      CALL "SENSOR CHECK" (
           Bit                      := "B 7.4",
           Preset_ms                := 500,
           Plc_Scan_ms              := "DB UTILITY".Scan_Cycle_Previous,
           Rising_Pulse_1           := "DB SENSOR CHECK".B7_4.Rising_Pulse_1,
           Rising_Pulse_2           := "DB SENSOR CHECK".B7_4.Rising_Pulse_2,
           Memory_Bit_1             := "DB SENSOR CHECK".B7_4.Memory_Bit_1,
           Memory_Bit_2             := "DB SENSOR CHECK".B7_4.Memory_Bit_2,
           Word_Buffer              := "DB SENSOR CHECK".B7_4.Word_buffer,
           Word_Result              := "DB SENSOR CHECK".B7_4.Word_Result);

NETWORK
TITLE =
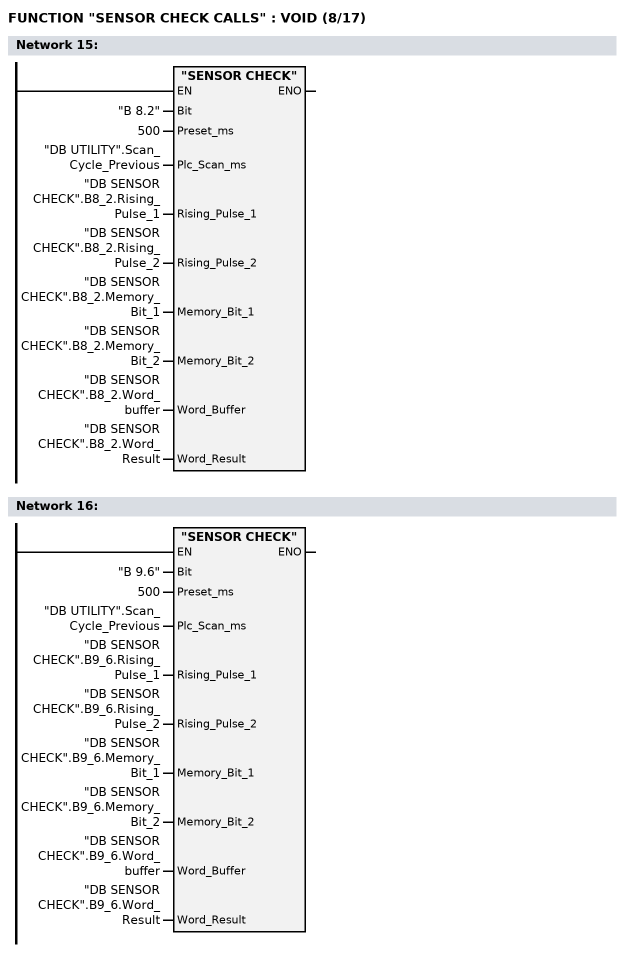

      CALL "SENSOR CHECK" (
           Bit                      := "B 8.2",
           Preset_ms                := 500,
           Plc_Scan_ms              := "DB UTILITY".Scan_Cycle_Previous,
           Rising_Pulse_1           := "DB SENSOR CHECK".B8_2.Rising_Pulse_1,
           Rising_Pulse_2           := "DB SENSOR CHECK".B8_2.Rising_Pulse_2,
           Memory_Bit_1             := "DB SENSOR CHECK".B8_2.Memory_Bit_1,
           Memory_Bit_2             := "DB SENSOR CHECK".B8_2.Memory_Bit_2,
           Word_Buffer              := "DB SENSOR CHECK".B8_2.Word_buffer,
           Word_Result              := "DB SENSOR CHECK".B8_2.Word_Result);

NETWORK
TITLE =

      CALL "SENSOR CHECK" (
           Bit                      := "B 9.6",
           Preset_ms                := 500,
           Plc_Scan_ms              := "DB UTILITY".Scan_Cycle_Previous,
           Rising_Pulse_1           := "DB SENSOR CHECK".B9_6.Rising_Pulse_1,
           Rising_Pulse_2           := "DB SENSOR CHECK".B9_6.Rising_Pulse_2,
           Memory_Bit_1             := "DB SENSOR CHECK".B9_6.Memory_Bit_1,
           Memory_Bit_2             := "DB SENSOR CHECK".B9_6.Memory_Bit_2,
           Word_Buffer              := "DB SENSOR CHECK".B9_6.Word_buffer,
           Word_Result              := "DB SENSOR CHECK".B9_6.Word_Result);

NETWORK
TITLE =
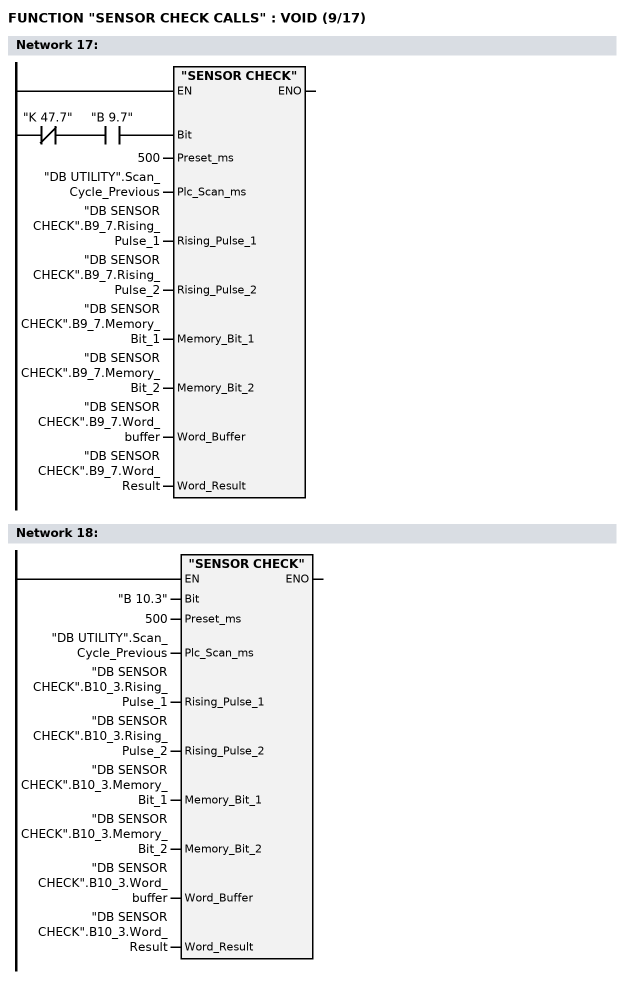

      AN    "K 47.7";
      A     "B 9.7";
      =     L      0.1;
//;
      CALL "SENSOR CHECK" (
           Bit                      := L      0.1,
           Preset_ms                := 500,
           Plc_Scan_ms              := "DB UTILITY".Scan_Cycle_Previous,
           Rising_Pulse_1           := "DB SENSOR CHECK".B9_7.Rising_Pulse_1,
           Rising_Pulse_2           := "DB SENSOR CHECK".B9_7.Rising_Pulse_2,
           Memory_Bit_1             := "DB SENSOR CHECK".B9_7.Memory_Bit_1,
           Memory_Bit_2             := "DB SENSOR CHECK".B9_7.Memory_Bit_2,
           Word_Buffer              := "DB SENSOR CHECK".B9_7.Word_buffer,
           Word_Result              := "DB SENSOR CHECK".B9_7.Word_Result);

NETWORK
TITLE =

      CALL "SENSOR CHECK" (
           Bit                      := "B 10.3",
           Preset_ms                := 500,
           Plc_Scan_ms              := "DB UTILITY".Scan_Cycle_Previous,
           Rising_Pulse_1           := "DB SENSOR CHECK".B10_3.Rising_Pulse_1,
           Rising_Pulse_2           := "DB SENSOR CHECK".B10_3.Rising_Pulse_2,
           Memory_Bit_1             := "DB SENSOR CHECK".B10_3.Memory_Bit_1,
           Memory_Bit_2             := "DB SENSOR CHECK".B10_3.Memory_Bit_2,
           Word_Buffer              := "DB SENSOR CHECK".B10_3.Word_buffer,
           Word_Result              := "DB SENSOR CHECK".B10_3.Word_Result);

NETWORK
TITLE =
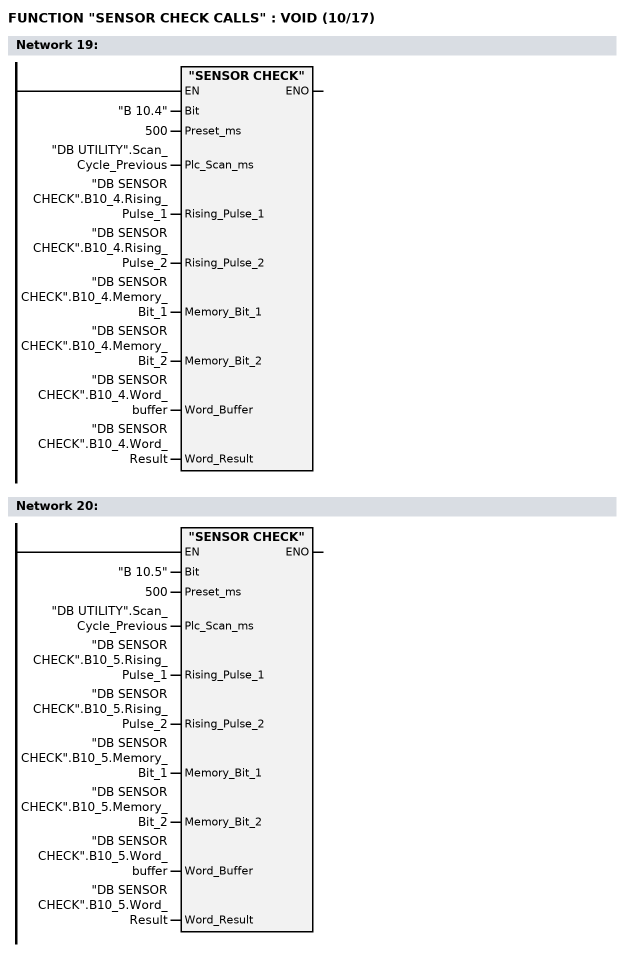

      CALL "SENSOR CHECK" (
           Bit                      := "B 10.4",
           Preset_ms                := 500,
           Plc_Scan_ms              := "DB UTILITY".Scan_Cycle_Previous,
           Rising_Pulse_1           := "DB SENSOR CHECK".B10_4.Rising_Pulse_1,
           Rising_Pulse_2           := "DB SENSOR CHECK".B10_4.Rising_Pulse_2,
           Memory_Bit_1             := "DB SENSOR CHECK".B10_4.Memory_Bit_1,
           Memory_Bit_2             := "DB SENSOR CHECK".B10_4.Memory_Bit_2,
           Word_Buffer              := "DB SENSOR CHECK".B10_4.Word_buffer,
           Word_Result              := "DB SENSOR CHECK".B10_4.Word_Result);

NETWORK
TITLE =

      CALL "SENSOR CHECK" (
           Bit                      := "B 10.5",
           Preset_ms                := 500,
           Plc_Scan_ms              := "DB UTILITY".Scan_Cycle_Previous,
           Rising_Pulse_1           := "DB SENSOR CHECK".B10_5.Rising_Pulse_1,
           Rising_Pulse_2           := "DB SENSOR CHECK".B10_5.Rising_Pulse_2,
           Memory_Bit_1             := "DB SENSOR CHECK".B10_5.Memory_Bit_1,
           Memory_Bit_2             := "DB SENSOR CHECK".B10_5.Memory_Bit_2,
           Word_Buffer              := "DB SENSOR CHECK".B10_5.Word_buffer,
           Word_Result              := "DB SENSOR CHECK".B10_5.Word_Result);

NETWORK
TITLE =
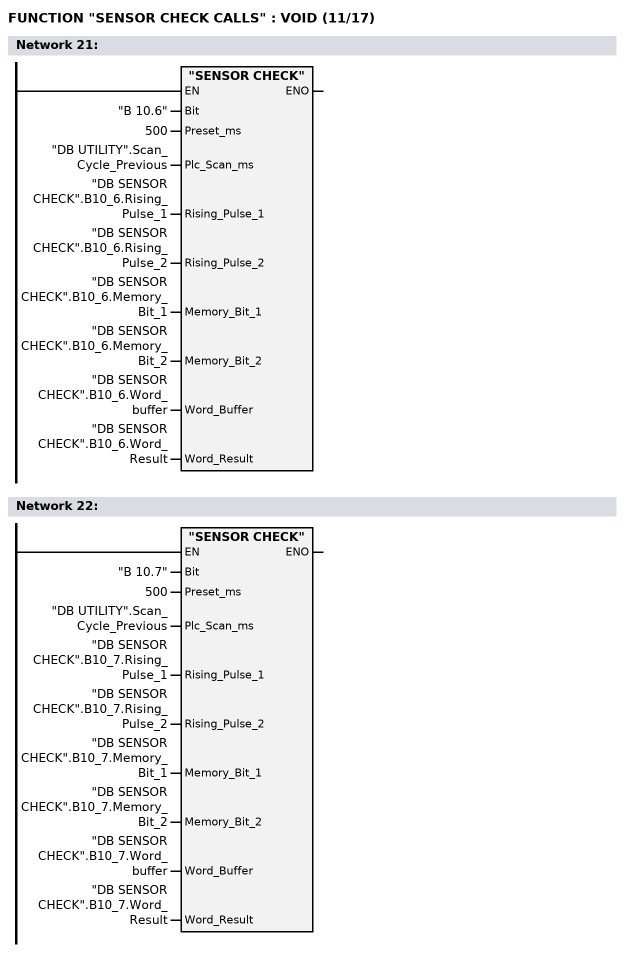

      CALL "SENSOR CHECK" (
           Bit                      := "B 10.6",
           Preset_ms                := 500,
           Plc_Scan_ms              := "DB UTILITY".Scan_Cycle_Previous,
           Rising_Pulse_1           := "DB SENSOR CHECK".B10_6.Rising_Pulse_1,
           Rising_Pulse_2           := "DB SENSOR CHECK".B10_6.Rising_Pulse_2,
           Memory_Bit_1             := "DB SENSOR CHECK".B10_6.Memory_Bit_1,
           Memory_Bit_2             := "DB SENSOR CHECK".B10_6.Memory_Bit_2,
           Word_Buffer              := "DB SENSOR CHECK".B10_6.Word_buffer,
           Word_Result              := "DB SENSOR CHECK".B10_6.Word_Result);

NETWORK
TITLE =

      CALL "SENSOR CHECK" (
           Bit                      := "B 10.7",
           Preset_ms                := 500,
           Plc_Scan_ms              := "DB UTILITY".Scan_Cycle_Previous,
           Rising_Pulse_1           := "DB SENSOR CHECK".B10_7.Rising_Pulse_1,
           Rising_Pulse_2           := "DB SENSOR CHECK".B10_7.Rising_Pulse_2,
           Memory_Bit_1             := "DB SENSOR CHECK".B10_7.Memory_Bit_1,
           Memory_Bit_2             := "DB SENSOR CHECK".B10_7.Memory_Bit_2,
           Word_Buffer              := "DB SENSOR CHECK".B10_7.Word_buffer,
           Word_Result              := "DB SENSOR CHECK".B10_7.Word_Result);

NETWORK
TITLE =
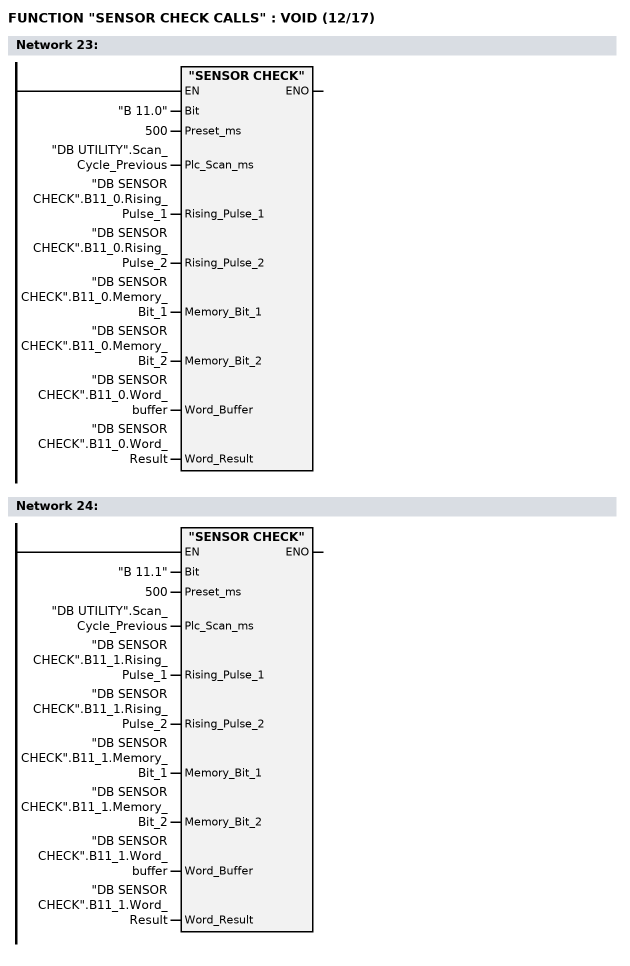

      CALL "SENSOR CHECK" (
           Bit                      := "B 11.0",
           Preset_ms                := 500,
           Plc_Scan_ms              := "DB UTILITY".Scan_Cycle_Previous,
           Rising_Pulse_1           := "DB SENSOR CHECK".B11_0.Rising_Pulse_1,
           Rising_Pulse_2           := "DB SENSOR CHECK".B11_0.Rising_Pulse_2,
           Memory_Bit_1             := "DB SENSOR CHECK".B11_0.Memory_Bit_1,
           Memory_Bit_2             := "DB SENSOR CHECK".B11_0.Memory_Bit_2,
           Word_Buffer              := "DB SENSOR CHECK".B11_0.Word_buffer,
           Word_Result              := "DB SENSOR CHECK".B11_0.Word_Result);

NETWORK
TITLE =

      CALL "SENSOR CHECK" (
           Bit                      := "B 11.1",
           Preset_ms                := 500,
           Plc_Scan_ms              := "DB UTILITY".Scan_Cycle_Previous,
           Rising_Pulse_1           := "DB SENSOR CHECK".B11_1.Rising_Pulse_1,
           Rising_Pulse_2           := "DB SENSOR CHECK".B11_1.Rising_Pulse_2,
           Memory_Bit_1             := "DB SENSOR CHECK".B11_1.Memory_Bit_1,
           Memory_Bit_2             := "DB SENSOR CHECK".B11_1.Memory_Bit_2,
           Word_Buffer              := "DB SENSOR CHECK".B11_1.Word_buffer,
           Word_Result              := "DB SENSOR CHECK".B11_1.Word_Result);

NETWORK
TITLE =
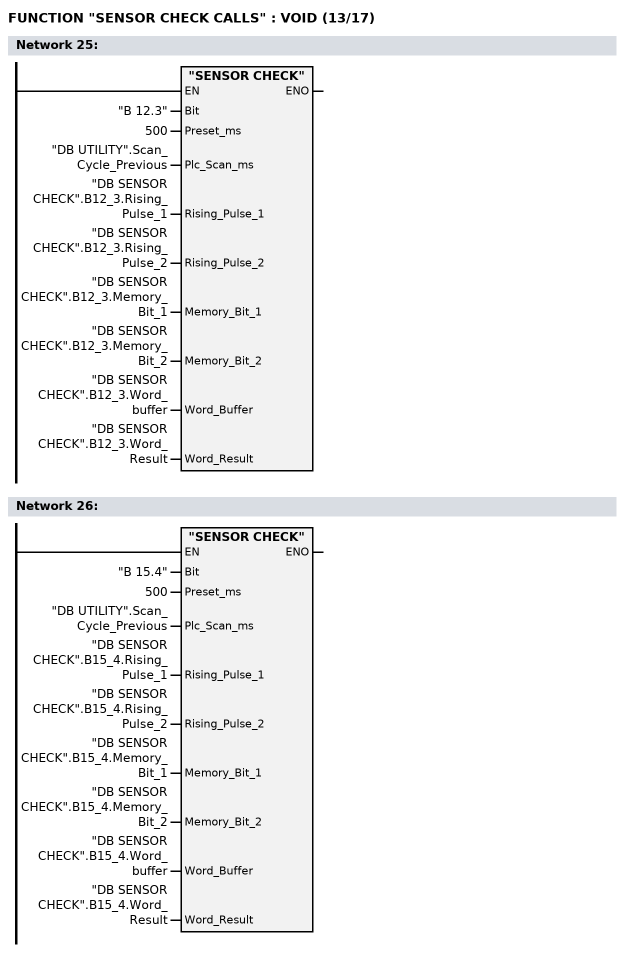

      CALL "SENSOR CHECK" (
           Bit                      := "B 12.3",
           Preset_ms                := 500,
           Plc_Scan_ms              := "DB UTILITY".Scan_Cycle_Previous,
           Rising_Pulse_1           := "DB SENSOR CHECK".B12_3.Rising_Pulse_1,
           Rising_Pulse_2           := "DB SENSOR CHECK".B12_3.Rising_Pulse_2,
           Memory_Bit_1             := "DB SENSOR CHECK".B12_3.Memory_Bit_1,
           Memory_Bit_2             := "DB SENSOR CHECK".B12_3.Memory_Bit_2,
           Word_Buffer              := "DB SENSOR CHECK".B12_3.Word_buffer,
           Word_Result              := "DB SENSOR CHECK".B12_3.Word_Result);

NETWORK
TITLE =

      CALL "SENSOR CHECK" (
           Bit                      := "B 15.4",
           Preset_ms                := 500,
           Plc_Scan_ms              := "DB UTILITY".Scan_Cycle_Previous,
           Rising_Pulse_1           := "DB SENSOR CHECK".B15_4.Rising_Pulse_1,
           Rising_Pulse_2           := "DB SENSOR CHECK".B15_4.Rising_Pulse_2,
           Memory_Bit_1             := "DB SENSOR CHECK".B15_4.Memory_Bit_1,
           Memory_Bit_2             := "DB SENSOR CHECK".B15_4.Memory_Bit_2,
           Word_Buffer              := "DB SENSOR CHECK".B15_4.Word_buffer,
           Word_Result              := "DB SENSOR CHECK".B15_4.Word_Result);

NETWORK
TITLE =
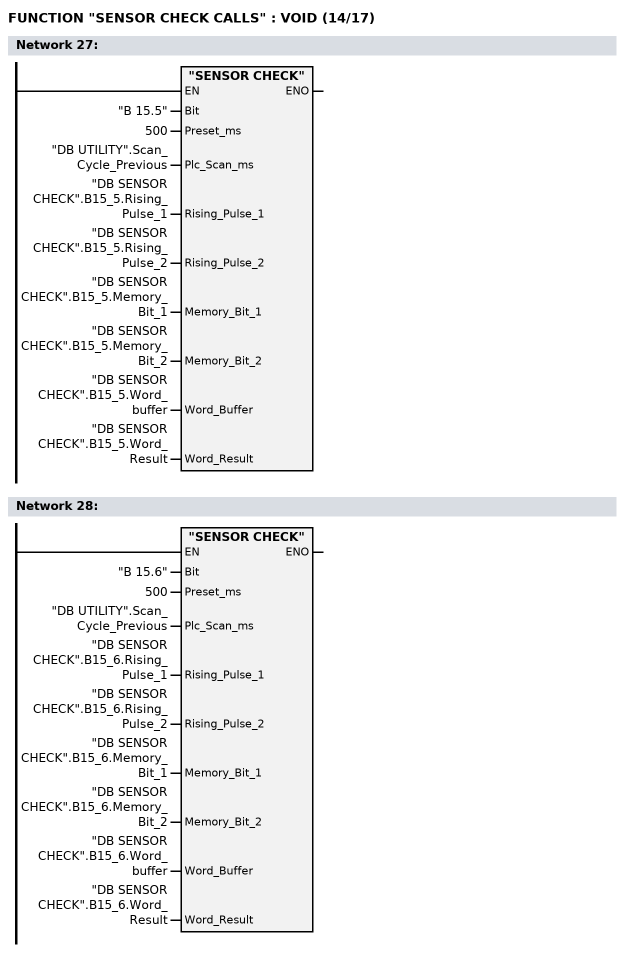

      CALL "SENSOR CHECK" (
           Bit                      := "B 15.5",
           Preset_ms                := 500,
           Plc_Scan_ms              := "DB UTILITY".Scan_Cycle_Previous,
           Rising_Pulse_1           := "DB SENSOR CHECK".B15_5.Rising_Pulse_1,
           Rising_Pulse_2           := "DB SENSOR CHECK".B15_5.Rising_Pulse_2,
           Memory_Bit_1             := "DB SENSOR CHECK".B15_5.Memory_Bit_1,
           Memory_Bit_2             := "DB SENSOR CHECK".B15_5.Memory_Bit_2,
           Word_Buffer              := "DB SENSOR CHECK".B15_5.Word_buffer,
           Word_Result              := "DB SENSOR CHECK".B15_5.Word_Result);

NETWORK
TITLE =

      CALL "SENSOR CHECK" (
           Bit                      := "B 15.6",
           Preset_ms                := 500,
           Plc_Scan_ms              := "DB UTILITY".Scan_Cycle_Previous,
           Rising_Pulse_1           := "DB SENSOR CHECK".B15_6.Rising_Pulse_1,
           Rising_Pulse_2           := "DB SENSOR CHECK".B15_6.Rising_Pulse_2,
           Memory_Bit_1             := "DB SENSOR CHECK".B15_6.Memory_Bit_1,
           Memory_Bit_2             := "DB SENSOR CHECK".B15_6.Memory_Bit_2,
           Word_Buffer              := "DB SENSOR CHECK".B15_6.Word_buffer,
           Word_Result              := "DB SENSOR CHECK".B15_6.Word_Result);

NETWORK
TITLE =
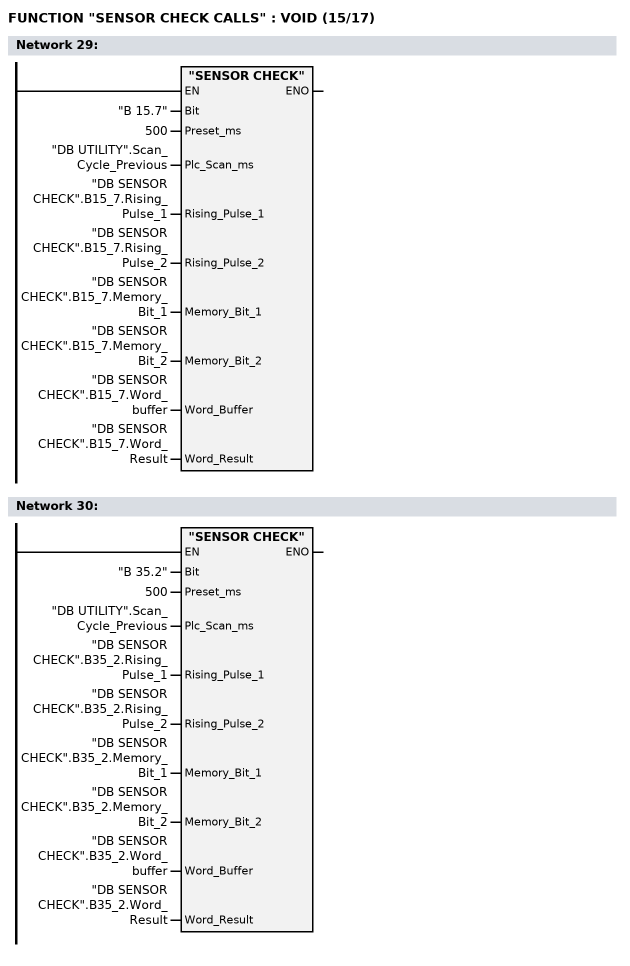

      CALL "SENSOR CHECK" (
           Bit                      := "B 15.7",
           Preset_ms                := 500,
           Plc_Scan_ms              := "DB UTILITY".Scan_Cycle_Previous,
           Rising_Pulse_1           := "DB SENSOR CHECK".B15_7.Rising_Pulse_1,
           Rising_Pulse_2           := "DB SENSOR CHECK".B15_7.Rising_Pulse_2,
           Memory_Bit_1             := "DB SENSOR CHECK".B15_7.Memory_Bit_1,
           Memory_Bit_2             := "DB SENSOR CHECK".B15_7.Memory_Bit_2,
           Word_Buffer              := "DB SENSOR CHECK".B15_7.Word_buffer,
           Word_Result              := "DB SENSOR CHECK".B15_7.Word_Result);

NETWORK
TITLE =

      CALL "SENSOR CHECK" (
           Bit                      := "B 35.2",
           Preset_ms                := 500,
           Plc_Scan_ms              := "DB UTILITY".Scan_Cycle_Previous,
           Rising_Pulse_1           := "DB SENSOR CHECK".B35_2.Rising_Pulse_1,
           Rising_Pulse_2           := "DB SENSOR CHECK".B35_2.Rising_Pulse_2,
           Memory_Bit_1             := "DB SENSOR CHECK".B35_2.Memory_Bit_1,
           Memory_Bit_2             := "DB SENSOR CHECK".B35_2.Memory_Bit_2,
           Word_Buffer              := "DB SENSOR CHECK".B35_2.Word_buffer,
           Word_Result              := "DB SENSOR CHECK".B35_2.Word_Result);

NETWORK
TITLE =
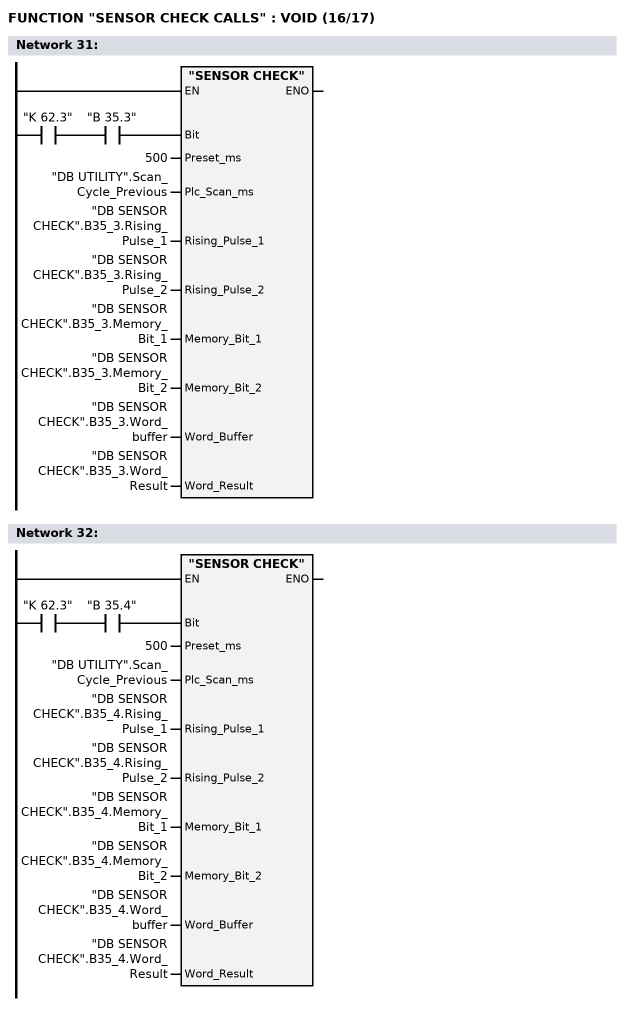

      A     "K 62.3";
      A     "B 35.3";
      =     L      0.2;

      CALL "SENSOR CHECK" (
           Bit                      := L      0.2,
           Preset_ms                := 500,
           Plc_Scan_ms              := "DB UTILITY".Scan_Cycle_Previous,
           Rising_Pulse_1           := "DB SENSOR CHECK".B35_3.Rising_Pulse_1,
           Rising_Pulse_2           := "DB SENSOR CHECK".B35_3.Rising_Pulse_2,
           Memory_Bit_1             := "DB SENSOR CHECK".B35_3.Memory_Bit_1,
           Memory_Bit_2             := "DB SENSOR CHECK".B35_3.Memory_Bit_2,
           Word_Buffer              := "DB SENSOR CHECK".B35_3.Word_buffer,
           Word_Result              := "DB SENSOR CHECK".B35_3.Word_Result);

NETWORK
TITLE =

      A     "K 62.3";
      A     "B 35.4";
      =     L      0.3;
//;
      CALL "SENSOR CHECK" (
           Bit                      := L      0.3,
           Preset_ms                := 500,
           Plc_Scan_ms              := "DB UTILITY".Scan_Cycle_Previous,
           Rising_Pulse_1           := "DB SENSOR CHECK".B35_4.Rising_Pulse_1,
           Rising_Pulse_2           := "DB SENSOR CHECK".B35_4.Rising_Pulse_2,
           Memory_Bit_1             := "DB SENSOR CHECK".B35_4.Memory_Bit_1,
           Memory_Bit_2             := "DB SENSOR CHECK".B35_4.Memory_Bit_2,
           Word_Buffer              := "DB SENSOR CHECK".B35_4.Word_buffer,
           Word_Result              := "DB SENSOR CHECK".B35_4.Word_Result);

NETWORK
TITLE =
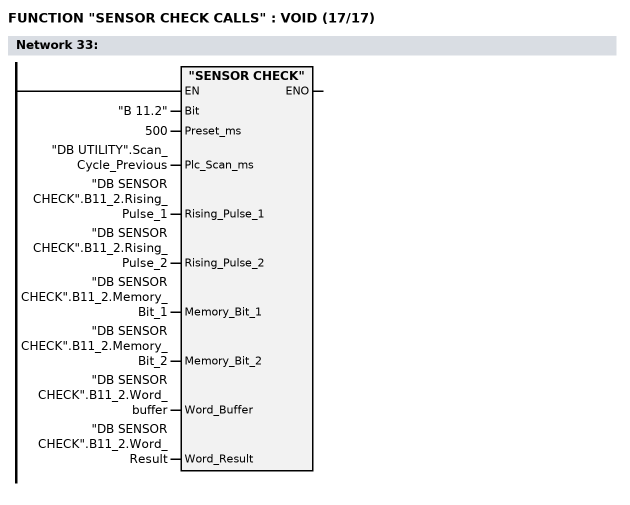

      CALL "SENSOR CHECK" (
           Bit                      := "B 11.2",
           Preset_ms                := 500,
           Plc_Scan_ms              := "DB UTILITY".Scan_Cycle_Previous,
           Rising_Pulse_1           := "DB SENSOR CHECK".B11_2.Rising_Pulse_1,
           Rising_Pulse_2           := "DB SENSOR CHECK".B11_2.Rising_Pulse_2,
           Memory_Bit_1             := "DB SENSOR CHECK".B11_2.Memory_Bit_1,
           Memory_Bit_2             := "DB SENSOR CHECK".B11_2.Memory_Bit_2,
           Word_Buffer              := "DB SENSOR CHECK".B11_2.Word_buffer,
           Word_Result              := "DB SENSOR CHECK".B11_2.Word_Result);

END_FUNCTION

FUNCTION "LAUER_RE-START_PUP" : VOID
TITLE =
//Logique de remise à zéro du bit de redémarrage de la communication avec
//l'interface.
//
//Ce bit doit être remis à zéro en cas de perte de communication avec l'automate
//ou si l'interface est éteint.
VERSION : 0.1

BEGIN
NETWORK
TITLE =Lauer restart bit
//DB50.DBW25 = S and mS   “Start a 5-second watchdog timer unless reset is
//active”
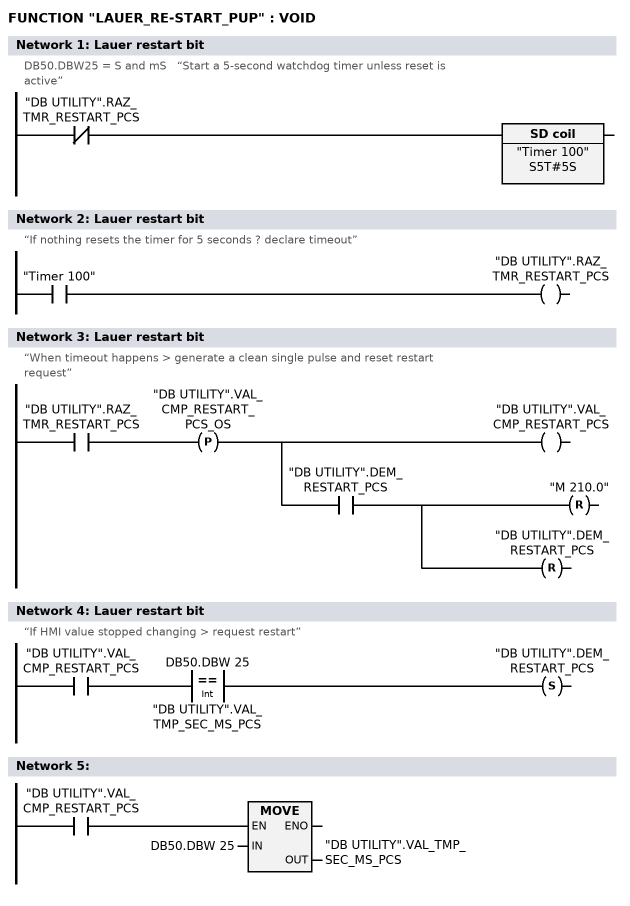
      AN    "DB UTILITY".RAZ_TMR_RESTART_PCS;
      L     S5T#5S;
      SD    "Timer 100";
      NOP   0;
      NOP   0;
      NOP   0;
      NOP   0;
NETWORK
TITLE =Lauer restart bit
//“If nothing resets the timer for 5 seconds ? declare timeout”
      A     "Timer 100";
      =     "DB UTILITY".RAZ_TMR_RESTART_PCS;
NETWORK
TITLE =Lauer restart bit
//“When timeout happens > generate a clean single pulse and reset restart
//request”
      A     "DB UTILITY".RAZ_TMR_RESTART_PCS;
      FP    "DB UTILITY".VAL_CMP_RESTART_PCS_OS;
      =     L      0.0;
      A     L      0.0;
      BLD   102;
      =     "DB UTILITY".VAL_CMP_RESTART_PCS;
      A     L      0.0;
      A     "DB UTILITY".DEM_RESTART_PCS;
      R     "M 210.0";
      R     "DB UTILITY".DEM_RESTART_PCS;
NETWORK
TITLE =Lauer restart bit
//“If HMI value stopped changing > request restart”
      A     "DB UTILITY".VAL_CMP_RESTART_PCS;
      A(    ;
      L     DB50.DBW   25;
      L     "DB UTILITY".VAL_TMP_SEC_MS_PCS;
      ==I   ;
      )     ;
      S     "DB UTILITY".DEM_RESTART_PCS;
NETWORK
TITLE =

      A     "DB UTILITY".VAL_CMP_RESTART_PCS;
      JNB   _001;
      L     DB50.DBW   25;
      T     "DB UTILITY".VAL_TMP_SEC_MS_PCS;
_001: NOP   0;
END_FUNCTION

FUNCTION "LAUER COMM ERR FC" : VOID
TITLE =
VERSION : 0.1

BEGIN
NETWORK
TITLE =
//;    Please choose your PCS and add the commands to your network
//;                      // Example PCS900/PCS 920/PCS950
//;                      // Typical presets
//;L W#16#1F00;  //(3F00 PCS950/PCS 920)
//;T DBW 72;
//;L W#16#00FF;
//;T DBW 74;
//;L W#16#0080;
//:T DBW 76;
//;                      // Example PCS009/PCS090/PCS095
//;                      // Typical presets
//;     L W#16#0FC8;
//;     T DBW 26;
//;     L W#16#0080;
//;     T DBW 28;
      L     W#16#0;
      T     DBW    8;
      T     DBW   10;
      T     DBW   12;
      T     DBW   14;
      T     DBW   46;
END_FUNCTION

FUNCTION "LAUER RESTART FC" : VOID
TITLE =
NAME : COFF
VERSION : 0.0

BEGIN
NETWORK
TITLE =
//;                     // Presets emergancy case
//;// Clear all keys
      L     W#16#0;
      T     DBW    8;
      T     DBW   10;
      T     DBW   12;
      T     DBW   14;
      T     DBW   46;
END_FUNCTION

FUNCTION "LAUER COMM FC" : VOID
TITLE =Handling Block Profibus
//
NAME : PROFIBUS
VERSION : 0.0


VAR_INPUT
  UBDB : BLOCK_DB ;	// UBDB
  RXFA : INT ;	// RXFA
  RXLE : INT ;	// RXLE
  TXFA : INT ;	// TXFA
  TXLE : INT ;	// TXLE
  RSET : BOOL ;	// RSET
  TIMT : TIMER ;	// TIMT
  TIMZ : S5TIME ;	// TIMZ
  COFF : BLOCK_FC ;	// COFF
  INIT : BLOCK_FC ;	// INIT
END_VAR
VAR_OUTPUT
  RFLM : BOOL ;	// RFLM
  EROR : BOOL ;	// EROR
END_VAR
VAR_TEMP
  conv_akku1 : DWORD ;
  conv_akku2 : DWORD ;
  conv_stw : WORD ;
END_VAR
BEGIN
NETWORK
TITLE =

      OPN   #UBDB; //  --------------------------
      AN    #RFLM; //  First action in FB?
      JC    OK;
      A     #TIMT; //  Timeout and no restart?
      AN    #RSET;
      JC    ERR;
      A     #TIMT;
      AN    #EROR;
      JC    ERR;
      JU    OK;

ERR:  A     #EROR;
      JC    ERR1;
      UC    #COFF; //  Call COFF once.
      OPN   #UBDB;

ERR1: A     #TIMT; //  If timeout set error-flag.
      S     #EROR;
      BEU   ;

OK:   A     #RFLM; //  First action?
      JC    CONT;
      UC    #INIT; //  Call INIT once.
      OPN   #UBDB;
      L     W#16#0; //  Init ----------------------
      T     DBW    0;
      T     DBW    2;
      T     DBW    4;
      T     DBW    6;
      AN    #RFLM;
      S     #RFLM; //  Set reset-ready-flag
//;
      AN    #RFLM; //  Trigger timer
      L     #TIMZ;
      SD    #TIMT;
//;
      A     #RFLM;
      L     #TIMZ;
      SD    #TIMT;

CONT: L     #RXFA;
      T     "MW 244"; //  ----------------------------
      +     1; //  Adress Handle1 E-Box
      T     "MW 252";
      L     #RXLE; //  Adress of first instruction
      +     -2;
      T     "MW 250"; //  Lenght E-Box Userdatas
//;
      L     #TXFA;
      T     "MW 242";
      +     1; //  Adress Handle1 A-Box
      T     "MW 248";
      L     #TXLE; //  Adress of first senddata
      +     -2;
      T     "MW 246"; //  Lenght A-Box-Userdatas
//;
      L     "MW 244"; //  Handle2 != Handle1? ---------
      L     #RXLE;
      +I    ;
      +     -1;
      T     "MW 238"; //  Adress Handle2
      T     #conv_akku1;
//;
      L     STW;
      T     #conv_stw;
//;
      L     "MB 239";
      SLW   3;
      LAR1  ;
      L     #conv_stw;
      T     STW;
//;
      L     #conv_akku1;
      L     IB [AR1,P#0.0];
      T     "MW 238"; //  Handle2
      T     #conv_akku1; //  Adress Handle1
//;
      L     STW;
      T     #conv_stw;
//;
      L     "MB 245";
      SLW   3;
      LAR1  ;
      L     #conv_stw;
      T     STW;
//;
      L     #conv_akku1;
      L     IB [AR1,P#0.0];
      L     "MW 238";
      <>I   ;
      BEC   ; //  Handle1 != Handle2 -> EXIT
//;
      T     #conv_akku1; //  Handle1 != HandleAlt? -------

      L     STW;
      T     #conv_stw;
//;
      L     "MB 245";
      SLW   3;
      LAR1  ;
      L     #conv_stw;
      T     STW;
//;
      L     #conv_akku1;
      L     IB [AR1,P#0.0];
      L     DBW    0; //  HandleAlt in UBDB (0)
      ==I   ;
      BEC   ;
//;
      AN    #RFLM; //  Start timeout-timer
      L     #TIMZ;
      SD    #TIMT;
//;
      A     #RFLM;
      L     #TIMZ;
      SD    #TIMT;
//;
      T     #conv_akku1; //  First action requiered?
      L     STW;
      T     #conv_stw;
      L     "MB 245";
      SLW   3;
      LAR1  ;
      L     #conv_stw;
      T     STW;
//;
      L     #conv_akku1;
      L     IB [AR1,P#0.0];
      L     W#16#80; //  Handle == 0x80?
      <>I   ;
      JC    SLP1;
      A     #RSET; // Clear Restart-Flag.
      R     #RSET;

END:  NOP   0;

      T     #conv_akku1; // Get Handle1(E) from RX-Box.

      L     STW;
      T     #conv_stw;
//;
      L     "MB 245";
      SLW   3;
      LAR1  ;
      L     #conv_stw;
      T     STW;
//;
      L     #conv_akku1;
      L     IB [AR1,P#0.0];
      T     DBW    0; // Save to HandleAlt.
      INVI  ; // Invert.
      T     "MW 236"; // Temporary saved.
      L     "MW 236";
      T     #conv_akku1; // Take inverted Handle1(E) to
      TAK   ;
      T     #conv_akku2;
      L     STW;
      T     #conv_stw;
//;
      L     "MB 243";
      SLW   3;
      LAR1  ;
      L     #conv_stw;
      T     STW;
//;
      L     #conv_akku2;
      L     #conv_akku1;
      T     QB [AR1,P#0.0]; // Handle1(A).
//;
      L     "MW 242";
      L     #TXLE;
      +I    ;
      +     -1;
      T     "MW 238"; // Take inverted Handle1(E) to
      L     "MW 236";
      T     #conv_akku1;
      TAK   ;
      T     #conv_akku2;
      L     STW;
      T     #conv_stw;
//;
      L     "MB 239";
      SLW   3;
      LAR1  ;
      L     #conv_stw;
      T     STW;
//;
      L     #conv_akku2;
      L     #conv_akku1;
      T     QB [AR1,P#0.0];
//;
      AN    #TIMT; // Clear Error-Mark.
      R     #EROR;
      BEU   ; // see you later...

SLP1: L     #RXFA; // Reached Rx-Box-End?
      L     #RXLE;
      +I    ;
      +     -1;
      L     "MW 252";
      ==I   ;
      JC    END;

      T     #conv_akku1; //  Start/Continue--------------

      L     STW;
      T     #conv_stw;
//;
      L     "MB 253";
      SLW   3;
      LAR1  ;
      L     #conv_stw;
      T     STW;
//;
      L     #conv_akku1;
      L     IW [AR1,P#0.0];
      L     W#16#0; //  Is anything usable?
      ==I   ;
      JC    END;

      T     #conv_akku1; //  Get first ABW.

      L     STW;
      T     #conv_stw;
//;
      L     "MB 253";
      SLW   3;
      LAR1  ;
      L     #conv_stw;
      T     STW;
//;
      L     #conv_akku1;
      L     IB [AR1,P#0.0];
      T     "MW 240"; //  Adress(UBDB) in ABW.
      L     "MW 252";
      +     1; //  Increment RX-Pointer.
      T     "MW 252";
      T     #conv_akku1;
      L     STW;
      T     #conv_stw;
      L     "MB 253";
      SLW   3;
      LAR1  ;
      L     #conv_stw;
      T     STW;
//;
      L     #conv_akku1;
      L     IB [AR1,P#0.0]; //  Count of ABW: Bit3..0.
      T     "MW 238"; //  Command of ABW: Bit 7..4.
      L     "MW 252"; //  ABW pointer to next ABW
      +     1; //  or first data.
      T     "MW 252";
//;
      L     "MW 238"; //  Check for right command.
      L     W#16#F0;
      AW    ;
      T     "MW 236"; //  Temporary saved.
//;
      L     "MW 236";
      L     W#16#10;
      ==I   ;
      JC    IOK;
//;
      L     "MW 236";
      L     W#16#20;
      ==I   ;
      JC    IOK;
//;
      L     "MW 236";
      L     W#16#40;
      ==I   ;
      JC    IOK;
//;
      L     "MW 236";
      L     W#16#80;
      ==I   ;
      JC    IOK;
      BEU   ; //  Command is wrong!
//;
IOK:  L     "MW 238"; //  Command is ok.
SLP2: L     W#16#F;
      AW    ; //  Count == 0:
      JZ    SLP1; //  Next subpaket
//;
      AN    "M 239.4";
      JC    ELS1;
      OPN   #UBDB;

      T     #conv_akku1; //  Offset ABW Adress in UBDB

      L     STW;
      T     #conv_stw;
//;
      L     "MB 241";
      SLW   4;
      LAR1  ;
      L     #conv_stw;
      T     STW;
//;
      L     #conv_akku1;
      L     DBW [AR1,P#0.0];
      T     #conv_akku1; //  Pointer to TX-Box
      TAK   ;
      T     #conv_akku2;
      L     STW;
      T     #conv_stw;
//;
      L     "MB 249";
      SLW   3;
      LAR1  ;
      L     #conv_stw;
      T     STW;
//;
      L     #conv_akku2;
      L     #conv_akku1;
      T     QW [AR1,P#0.0]; //  Write to TX-Box.
      L     "MW 248";
      +     2;
      T     "MW 248";
      JU    COMM;

ELS1: NOP   0;

      T     #conv_akku1; //  Pointer to RX-Box.

      L     STW;
      T     #conv_stw;
//;
      L     "MB 253";
      SLW   3;
      LAR1  ;
      L     #conv_stw;
      T     STW;
//;
      L     #conv_akku1;
      L     IW [AR1,P#0.0];
      T     "MW 236"; //  Read Data/Mask from RX-Box.
      L     "MW 252"; //  Increment Pointer to RX-Box.
      +     2;
      T     "MW 252";
//;
      AN    "M 239.5"; //  WRITE/(AND/OR)
      JC    ELS2;
      L     "MW 236";
      OPN   #UBDB;

      T     #conv_akku1; //  Offset ABW Adress in UBDB.
      TAK   ;
      T     #conv_akku2;
      L     STW;
      T     #conv_stw;
      L     "MB 241";
      SLW   4;
      LAR1  ;
      L     #conv_stw;
      T     STW;
//;
      L     #conv_akku2;
      L     #conv_akku1;
      T     DBW [AR1,P#0.0]; //  Write to UBDB.
      JU    COMM;

ELS2: AN    "M 239.6";
      JC    ELS3;
      L     "MW 236";
      OPN   #UBDB;

      T     #conv_akku1; //  Offset ABW Adress in UBDB.
      L     STW;
      T     #conv_stw;
      L     "MB 241";
      SLW   4;
      LAR1  ;
      L     #conv_stw;
      T     STW;
//;
      L     #conv_akku1;
      L     DBW [AR1,P#0.0];
      AW    ;
      OPN   #UBDB;
      T     #conv_akku1;
      TAK   ;
      T     #conv_akku2;
      L     STW;
      T     #conv_stw;
      L     "MB 241";
      SLW   4;
      LAR1  ;
      L     #conv_stw;
      T     STW;
//;
      L     #conv_akku2;
      L     #conv_akku1;
      T     DBW [AR1,P#0.0]; //  And to UBDB
      JU    COMM;

ELS3: NOP   0;

      L     "MW 236";
      OPN   #UBDB;
      T     #conv_akku1;
      L     STW;
      T     #conv_stw;
      L     "MB 241";
      SLW   4;
      LAR1  ;
      L     #conv_stw;
      T     STW;
//;
      L     #conv_akku1;
      L     DBW [AR1,P#0.0];
      OW    ;
      OPN   #UBDB;

      T     #conv_akku1;
      TAK   ;
      T     #conv_akku2;
      L     STW;
      T     #conv_stw;
      L     "MB 241";
      SLW   4;
      LAR1  ;
      L     #conv_stw;
      T     STW;
//;
      L     #conv_akku2;
      L     #conv_akku1;
      T     DBW [AR1,P#0.0];
COMM: L     "MW 240";
      +     1;
      T     "MW 240";
      L     "MW 238"; //  Decrement counter of ABW.
      +     -1;
      T     "MW 238";
      JU    SLP2;
END_FUNCTION

FUNCTION "LAUER" : VOID
TITLE =
NAME : SCHRIANZ
VERSION : 0.0


VAR_TEMP
  TEMP0 : DWORD ;
  TEMP1 : DWORD ;
  TEMP2 : WORD ;
END_VAR
BEGIN
NETWORK
TITLE =



NETWORK
TITLE =



NETWORK
TITLE =

      OPN   "DB LAUER";

NETWORK
TITLE =

      AN    "M 150.7";
      JC    M001;
      L     2#100000000;
      T     DBW   72;
M001: NOP   0;
NETWORK
TITLE =

      ON    "M 150.7";
      JC    M002;
      L     2#1;
      T     DBW   76;
M002: NOP   0;
NETWORK
TITLE =



NETWORK
TITLE =

      O(    ;
      L     DBW  300;
      L     77;
      <I    ;
      )     ;
      O(    ;
      L     DBW  300;
      L     102;
      >I    ;
      )     ;
      JC    M003;
      JU    M004;
M003: L     77;
      T     DBW  300;
M004: NOP   0;
NETWORK
TITLE =

      L     "DB LAUER".D_150;
      L     77;
      <>I   ;
      JC    M005;
      L     "MW 15";
      T     "MW 200";
      L     "MB 17";
      T     MB   202;
M005: L     DBW  300;
      L     78;
      <>I   ;
      JC    M006;
      L     "MW 19";
      T     "MW 200";
      L     "MB 21";
      T     MB   202;
M006: L     DBW  300;
      L     79;
      <>I   ;
      JC    M007;
      L     "MW 23";
      T     "MW 200";
      L     "MB 25";
      T     MB   202;
M007: L     DBW  300;
      L     80;
      <>I   ;
      JC    M008;
      L     "MW 27";
      T     "MW 200";
      L     "MB 29";
      T     MB   202;
M008: L     DBW  300;
      L     81;
      <>I   ;
      JC    M009;
      L     "MW 31";
      T     "MW 200";
      L     "MB 33";
      T     MB   202;
M009: L     DBW  300;
      L     82;
      <>I   ;
      JC    M00a;
      L     "MW 35";
      T     "MW 200";
      L     "MB 37";
      T     MB   202;
M00a: L     DBW  300;
      L     83;
      <>I   ;
      JC    M00b;
      L     "MW 39";
      T     "MW 200";
      L     "MB 41";
      T     MB   202;
M00b: L     DBW  300;
      L     84;
      <>I   ;
      JC    M00c;
      L     "MW 43";
      T     "MW 200";
      L     "MB 45";
      T     MB   202;
M00c: L     DBW  300;
      L     85;
      <>I   ;
      JC    M00d;
      L     "MW 47";
      T     "MW 200";
      L     "MB 49";
      T     MB   202;
M00d: L     DBW  300;
      L     86;
      <>I   ;
      JC    M00e;
      L     "MW 51";
      T     "MW 200";
      L     "MB 53";
      T     MB   202;
M00e: L     DBW  300;
      L     87;
      <>I   ;
      JC    M00f;
      L     "MW 55";
      T     "MW 200";
      L     "MB 57";
      T     MB   202;
M00f: L     DBW  300;
      L     88;
      <>I   ;
      JC    M010;
      L     "MW 59";
      T     "MW 200";
      L     "MB 61";
      T     MB   202;
M010: L     DBW  300;
      L     89;
      <>I   ;
      JC    M011;
      L     "MW 63";
      T     "MW 200";
      T     "MW 200";
      L     "MB 65";
      T     MB   202;
M011: L     DBW  300;
      L     90;
      <>I   ;
      JC    M012;
      L     "MW 67";
      T     "MW 200";
      L     "MB 69";
      T     MB   202;
M012: L     DBW  300;
      L     91;
      <>I   ;
      JC    M013;
      L     "MW 71";
      T     "MW 200";
      L     "MB 73";
      T     MB   202;
M013: L     DBW  300;
      L     92;
      <>I   ;
      JC    M014;
      L     "MW 75";
      T     "MW 200";
      L     "MB 77";
      T     MB   202;
M014: L     DBW  300;
      L     93;
      <>I   ;
      JC    M015;
      L     "MW 79";
      T     "MW 200";
      L     "MB 81";
      T     MB   202;
M015: L     DBW  300;
      L     94;
      <>I   ;
      JC    M016;
      L     "MW 83";
      T     "MW 200";
      L     "MB 85";
      T     MB   202;
M016: L     DBW  300;
      L     95;
      <>I   ;
      JC    M017;
      L     "MW 87";
      T     "MW 200";
      L     "MB 89";
      T     MB   202;
M017: L     DBW  300;
      L     96;
      <>I   ;
      JC    M018;
      L     "MW 91";
      T     "MW 200";
      L     "MB 93";
      T     MB   202;
M018: L     DBW  300;
      L     97;
      <>I   ;
      JC    M019;
      L     "MW 95";
      T     "MW 200";
      L     "MB 97";
      T     MB   202;
M019: L     DBW  300;
      L     98;
      <>I   ;
      JC    M01a;
      L     "MW 99";
      T     "MW 200";
      L     "MB 101";
      T     MB   202;
M01a: L     DBW  300;
      L     99;
      <>I   ;
      JC    M01b;
      L     "MW 103";
      T     "MW 200";
      L     "MB 105";
      T     MB   202;
M01b: L     DBW  300;
      L     100;
      <>I   ;
      JC    M01c;
      L     "MW 107";
      T     "MW 200";
      L     "MB 109";
      T     MB   202;
M01c: L     DBW  300;
      L     101;
      <>I   ;
      JC    M01d;
      L     "MW 111";
      L     "MW 200";
      L     "MB 113";
      T     MB   202;
M01d: L     DBW  300;
      L     102;
      <>I   ;
      JC    M01e;
      L     "MW 115";
      T     "MW 200";
      L     "MB 117";
      T     MB   202;
M01e: NOP   0;
NETWORK
TITLE =

      L     W#16#0;
      T     MB   204;
      L     W#16#80;
      T     MB   207;
NETWORK
TITLE =

      AN    "M 203.0";
      JC    M01f;
      L     25;
      T     MB   204;
M020: L     MB   203;
      SRW   1;
      T     MB   203;
      L     MB   207;
      SRW   1;
      T     "MW 207";
      AN    "M 203.0";
      JC    M021;
      L     MB   204;
      INC   1;
      T     MB   204;
M021: AN    "M 207.0";
      JC    M020;
      JU    M022;
M01f: AN    "M 202.0";
      JC    M023;
      L     17;
      T     MB   204;
M024: L     MB   202;
      SRW   1;
      T     MB   202;
      L     MB   207;
      SRW   1;
      T     MB   207;
      AN    "M 202.0";
      JC    M025;
      L     MB   204;
      INC   1;
      T     MB   204;
M025: AN    "M 207.0";
      JC    M024;
      JU    M022;
M023: AN    "M 201.0";
      JC    M026;
      L     9;
      T     MB   204;
M027: L     "MB 201";
      SRW   1;
      T     "MB 201";
      L     MB   207;
      SRW   1;
      T     MB   207;
      AN    "M 201.0";
      JC    M028;
      L     MB   204;
      INC   1;
      T     MB   204;
M028: AN    "M 207.0";
      JC    M027;
      JU    M022;
M026: AN    "M 200.0";
      JC    M022;
      L     1;
      T     MB   204;
M029: L     "MB 200";
      SRW   1;
      T     "MB 200";
      L     MB   207;
      SRW   1;
      T     MB   207;
      AN    "M 200.0";
      JC    M02a;
      L     MB   204;
      INC   1;
      T     MB   204;
M02a: AN    "M 207.0";
      JC    M029;
M022: NOP   0;
NETWORK
TITLE =



NETWORK
TITLE =

      OPN   "DB LAUER";
      L     MB   204;
      T     #TEMP0;
      TAK   ;
      T     #TEMP1;
      L     STW;
      T     #TEMP2;
      L     DBB  301;
      SLW   4;
      LAR1  ;
      L     #TEMP2;
      T     STW;
      L     #TEMP1;
      L     #TEMP0;
      T     DBW [AR1,P#0.0];
NETWORK
TITLE =



NETWORK
TITLE =

      L     "DB LAUER".D_150;
      INC   1;
      T     DBW  300;
NETWORK
TITLE =



NETWORK
TITLE =



END_FUNCTION

FUNCTION "CONTROL" : VOID
TITLE =Controls
VERSION : 0.0

BEGIN
NETWORK
TITLE =Qty Accumulation Conveyor
//  A     "M 0.3"
//      A     "M 92.0"
//      AN    "M 14.4"
//      CU    "COUNTER 4"
////;
//      A     "M 0.3"
//      A     "B 6.4"
//      CD    "COUNTER 4"
////;
//      A     "M 161.0"
//      A     "M 161.1"
//      A(
//      ON    "S 2.1"
//      O     "S 2.2"
//      )
//      R     "COUNTER 4"
//


NETWORK
TITLE =Qty Accumulation Conveyor
//      A     "M 0.3"
//      AN    "B 6.7"
//      CU    "COUNTER 5"
//      A     "M 0.3"
//      AN    "B 7.2"
//      CD    "COUNTER 5"
//      A     "M 161.0"
//      A     "M 161.1"
//      A(
//      ON    "S 2.1"
//      O     "S 2.2"
//      )
//      R     "COUNTER 5"
//


NETWORK
TITLE =Qty Flipper to Pusher
//      A     "M 0.3"
//      AN    "B 7.4"
//      CU    "COUNTER 6"
//      A     "M 0.3"
//      AN    "B 10.4"
//      CD    "COUNTER 6"
//      A     "M 161.0"
//      A     "M 161.1"
//      A(
//      ON    "S 2.1"
//      O     "S 2.2"
//      )
//      R     "COUNTER 6"
//


NETWORK
TITLE =Qty Pivot / Collator Conveyor
//      A     "M 0.3"
//      AN    "B 10.4"
//      CU    "COUNTER 7"
//      A     "M 0.3"
//      AN    "B 10.5"
//      CD    "COUNTER 7"
//      A     "M 161.0"
//      A     "M 161.1"
//      A(
//      ON    "S 2.1"
//      O     "S 2.2"
//      )
//      R     "COUNTER 7"
//


NETWORK
TITLE =Qty Bottom Accumulator
//      A     "M 0.3"
//      A     "B 10.6"
//      A     "P 15.1"
//      CU    "COUNTER 8"
//      A     "M 0.3"
//      AN    "B 11.2"
//      CD    "COUNTER 8"
//      A     "M 161.0"
//      A     "M 161.1"
//      A(
//      ON    "S 2.1"
//      O     "S 2.2"
//      )
//      R     "COUNTER 8"
//


NETWORK
TITLE =Qty Top Accumulator
//      A     "M 0.3"
//      A     "B 10.6"
//      A     "P 15.0"
//      CU    "COUNTER 9"
//      A     "M 0.3"
//      AN    "B 15.6"
//      CD    "COUNTER 9"
//      A     "M 161.1"
//      A     "M 161.1"
//      A(
//      ON    "S 2.1"
//      O     "S 2.2"
//      )
//      R     "COUNTER 9"
//


NETWORK
TITLE =Start Signal
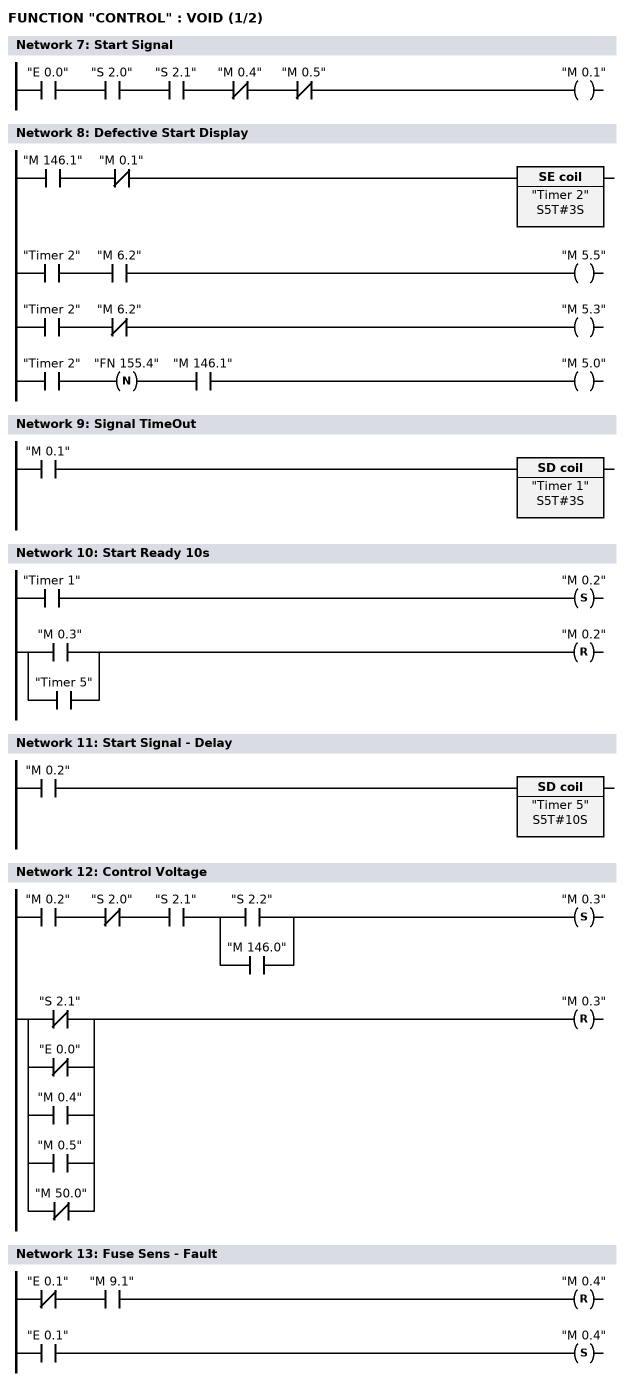

      A     "E 0.0";
      A(    ;
      O     "S 2.0";
//   O     "M 146.1"
      )     ;
      A     "S 2.1";
//      A     "M 146.2"
      AN    "M 0.4";
      AN    "M 0.5";
      =     "M 0.1";
NETWORK
TITLE =Defective Start Display

      A     "M 146.1";
      AN    "M 0.1";
      L     S5T#3S;
      SE    "Timer 2";
//;
      A     "Timer 2";
      A     "M 6.2";
      =     "M 5.5";
//;
      A     "Timer 2";
      AN    "M 6.2";
      =     "M 5.3";
//;
      A     "Timer 2";
      FN    "FN 155.4";
      A     "M 146.1";
      =     "M 5.0";
NETWORK
TITLE =Signal TimeOut

      A     "M 0.1";
      L     S5T#3S;
      SD    "Timer 1";
NETWORK
TITLE =Start Ready 10s

      A     "Timer 1";
      S     "M 0.2";
//;
      A(    ;
      O     "M 0.3";
      O     "Timer 5";
      )     ;
      R     "M 0.2";
NETWORK
TITLE =Start Signal - Delay

      A     "M 0.2";
      L     S5T#10S;
      SD    "Timer 5";
NETWORK
TITLE =Control Voltage

      A     "M 0.2";
      AN    "S 2.0";
      A     "S 2.1";
//    A    "M 146.2"
      A(    ;
      O     "S 2.2";
      O     "M 146.0";
      )     ;
      S     "M 0.3";
//;
      A(    ;
      ON    "S 2.1";
//    ON    "M 146.2"
      ON    "E 0.0";
      O     "M 0.4";
      O     "M 0.5";
      ON    "M 50.0";
      )     ;
      R     "M 0.3";
NETWORK
TITLE =Fuse Sens - Fault

      AN    "E 0.1";
      A     "M 9.1";
      R     "M 0.4";
//;
      A     "E 0.1";
      S     "M 0.4";
NETWORK
TITLE =Motor Protect - Fault
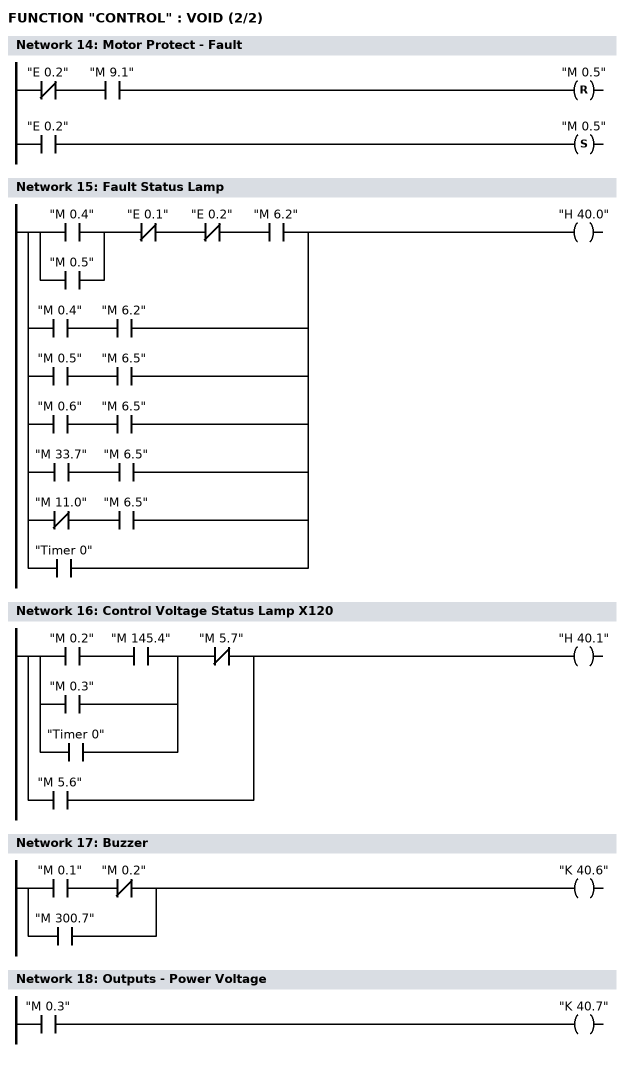

      AN    "E 0.2";
      A     "M 9.1";
      R     "M 0.5";
//;
      A     "E 0.2";
      S     "M 0.5";
NETWORK
TITLE =Fault Status Lamp

      A(    ;
      O     "M 0.4";
      O     "M 0.5";
      )     ;
      AN    "E 0.1";
      AN    "E 0.2";
      A     "M 6.2";
      O     ;
      A     "M 0.4";
      A     "M 6.2";
      O     ;
      A     "M 0.5";
      A     "M 6.5";
      O     ;
      A     "M 0.6";
      A     "M 6.5";
      O     ;
      A     "M 33.7";
      A     "M 6.5";
      O     ;
      AN    "M 11.0";
      A     "M 6.5";
      O     "Timer 0";
      =     "H 40.0";
NETWORK
TITLE =Control Voltage Status Lamp X120

      A     "M 0.2";
      A     "M 145.4";
      O     "M 0.3";
      O     "Timer 0";
      AN    "M 5.7";
      O     "M 5.6";
      =     "H 40.1";
NETWORK
TITLE =Buzzer

      A     "M 0.1";
      AN    "M 0.2";
      O     "M 300.7";
      =     "K 40.6";
NETWORK
TITLE =Outputs - Power Voltage

      A     "M 0.3";
      =     "K 40.7";
END_FUNCTION

FUNCTION "GENERAL FAULTS" : VOID
TITLE =General Faults
VERSION : 0.0


VAR_TEMP
  INIT_DELAY : BOOL ;
  CHECK_PULSE : BOOL ;
  ELEVATOR_U42_0 : BOOL ;	//CO ELEVATOR VFD U42.0 - READY    POS.2
  FAULT_TRIGGERED : BOOL ;
  FAULT_REGISTER_1 : BOOL ;
  FAULT_REGISTER_2 : BOOL ;
  FAULT_REGISTER_3 : BOOL ;
  FAULT_REGISTER_4 : BOOL ;
  FAULT_REGISTER_5 : BOOL ;
END_VAR
BEGIN
NETWORK
TITLE =Trigger Pulse
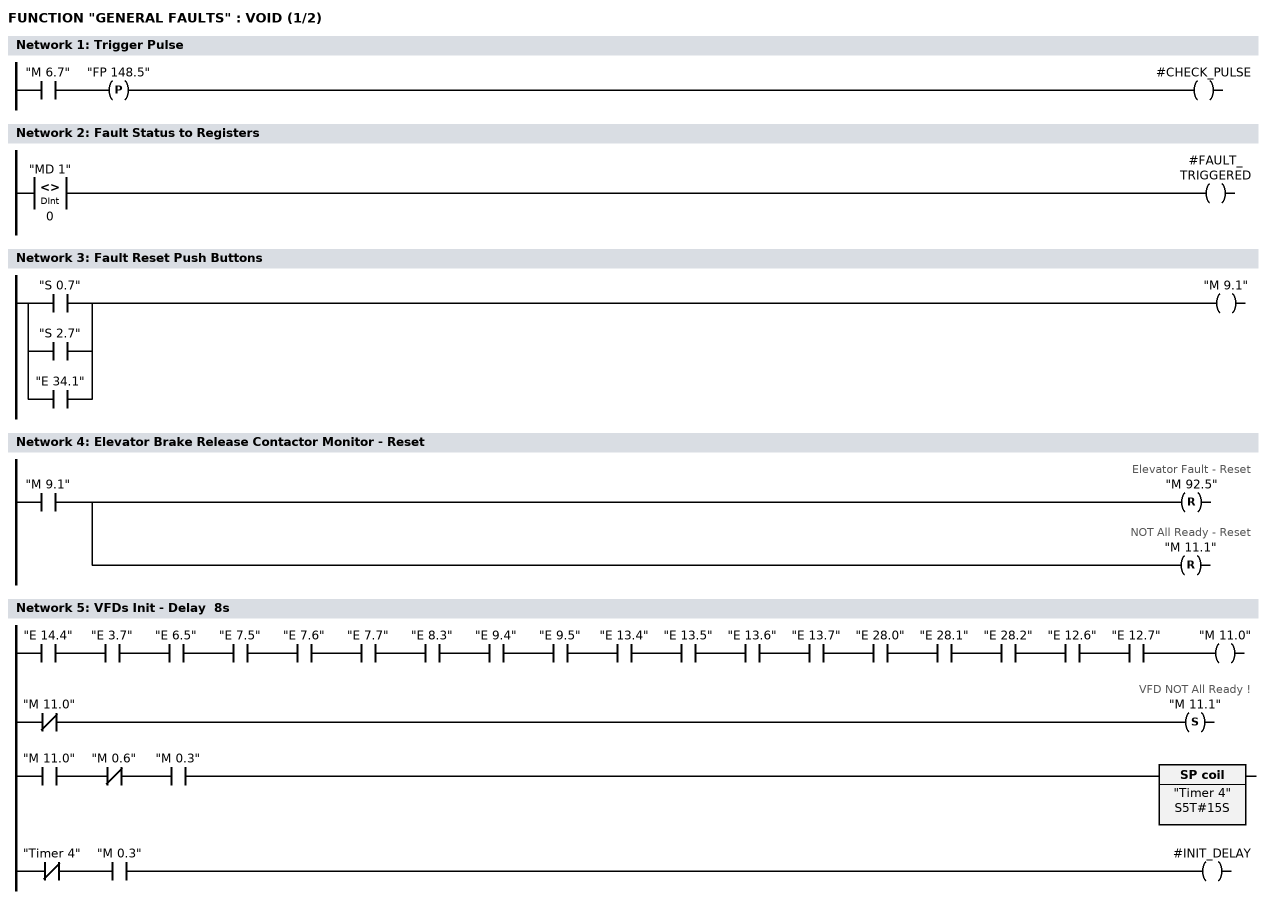

      A     "M 6.7";
      FP    "FP 148.5";
      =     #CHECK_PULSE;
NETWORK
TITLE =Fault Status to Registers

      A(    ;
      L     "MD 1";
      L     0;
      <>D   ;
      )     ;
      =     #FAULT_TRIGGERED;
NETWORK
TITLE =Fault Reset Push Buttons

      A(    ;
      O     "S 0.7";
      O     "S 2.7";
      O     "E 34.1";
      )     ;
      =     "M 9.1";
NETWORK
TITLE =Elevator Brake Release Contactor Monitor - Reset

      A     "M 9.1";
      R     "M 92.5"; // Elevator Fault - Reset
      R     "M 11.1"; // NOT All Ready - Reset
NETWORK
TITLE =VFDs Init - Delay  8s

      A(    ;
      A     "E 14.4";
      A     "E 3.7";
      A     "E 6.5";
      A     "E 7.5";
      A     "E 7.6";
      A     "E 7.7";
      A     "E 8.3";
      A     "E 9.4";
      A     "E 9.5";
      A     "E 13.4";
      A     "E 13.5";
      A     "E 13.6";
      A     "E 13.7";
      A     "E 28.0";
      A     "E 28.1";
      A     "E 28.2";
      A     "E 12.6";
      A     "E 12.7";
      )     ;
      =     "M 11.0";
//;
      AN    "M 11.0";
      S     "M 11.1"; // VFD NOT All Ready !
//;

      A     "M 11.0";
      AN    "M 0.6";
      A     "M 0.3";
      L     S5T#15S;
      SP    "Timer 4";
//;
      AN    "Timer 4";
      A     "M 0.3";
      =     #INIT_DELAY;
NETWORK
TITLE =Motor Temp Control - Fault Check
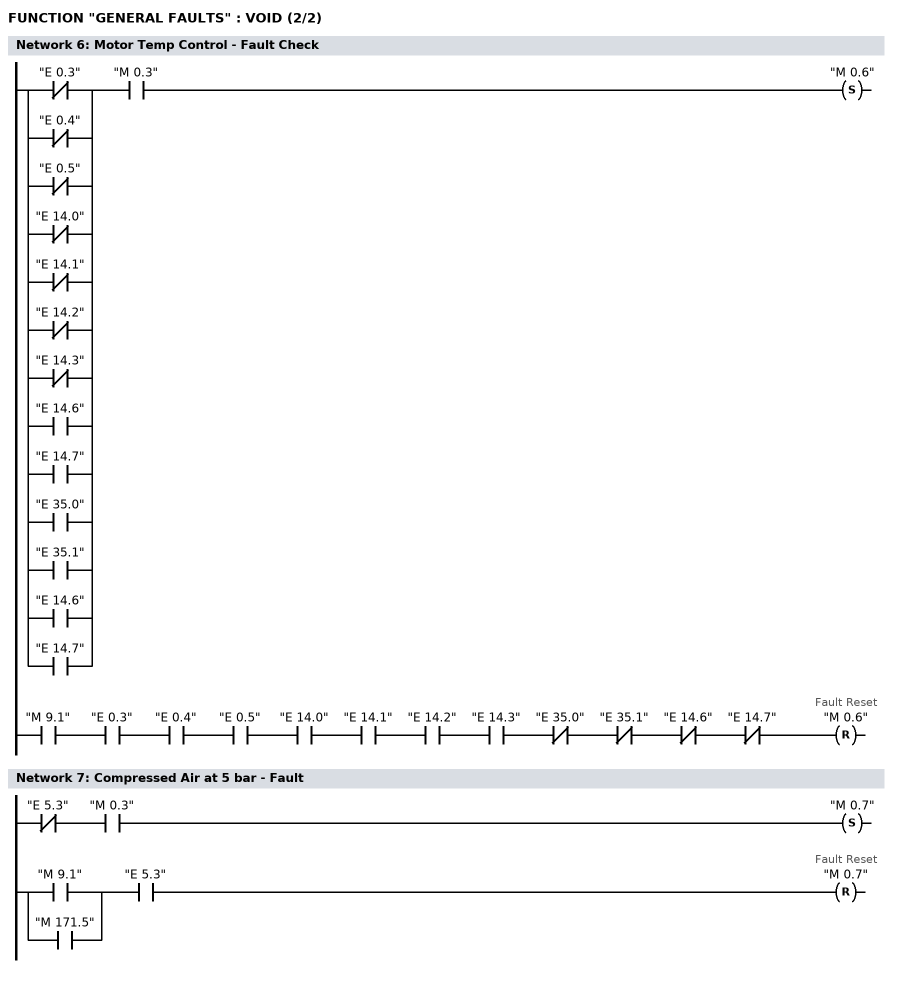

      A(    ;
      ON    "E 0.3";
      ON    "E 0.4";
      ON    "E 0.5";
      ON    "E 14.0";
      ON    "E 14.1";
      ON    "E 14.2";
      ON    "E 14.3";
      O     "E 14.6";
      O     "E 14.7";
      O     "E 35.0";
      O     "E 35.1";
      O     "E 14.6";
      O     "E 14.7";
      )     ;
      A     "M 0.3";
      S     "M 0.6";
//;
      A     "M 9.1";
      A     "E 0.3";
      A     "E 0.4";
      A     "E 0.5";
      A     "E 14.0";
      A     "E 14.1";
      A     "E 14.2";
      A     "E 14.3";
      AN    "E 35.0";
      AN    "E 35.1";
      AN    "E 14.6";
      AN    "E 14.7";
      R     "M 0.6"; // Fault Reset
NETWORK
TITLE =Compressed Air at 5 bar - Fault

      AN    "E 5.3";
      A     "M 0.3";
      S     "M 0.7";
//;
      A(    ;
      O     "M 9.1";
      O     "M 171.5";
      )     ;
      A     "E 5.3";
      R     "M 0.7"; // Fault Reset
NETWORK
TITLE =Faults Register 1 - E-Stops & Safety Doors

      A(    ;
      L     "MB 1";
      L     0;
      <>I   ;
      )     ;
      =     #FAULT_REGISTER_1;
//;
      A     #FAULT_REGISTER_1;
      O     #CHECK_PULSE;
      O     "M 17.1";
      O     "M 9.1";
      JNB   FR01;
NETWORK
TITLE =E-Stop  Desk  X120
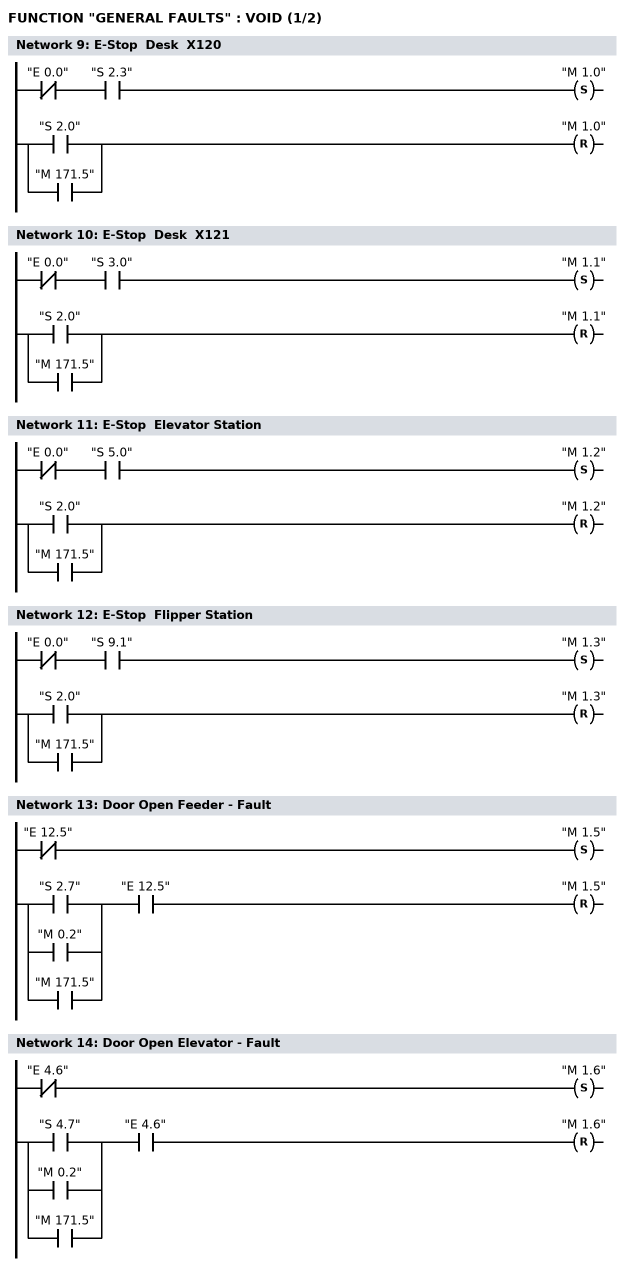

      AN    "E 0.0";
      A     "S 2.3";
      S     "M 1.0";
//;
      A(    ;
      O     "S 2.0";
      O     "M 171.5";
      )     ;
      R     "M 1.0";
NETWORK
TITLE =E-Stop  Desk  X121

      AN    "E 0.0";
      A     "S 3.0";
      S     "M 1.1";
//;
      A(    ;
      O     "S 2.0";
      O     "M 171.5";
      )     ;
      R     "M 1.1";
NETWORK
TITLE =E-Stop  Elevator Station

      AN    "E 0.0";
      A     "S 5.0";
      S     "M 1.2";
//;
      A(    ;
      O     "S 2.0";
      O     "M 171.5";
      )     ;
      R     "M 1.2";
NETWORK
TITLE =E-Stop  Flipper Station

      AN    "E 0.0";
      A     "S 9.1";
      S     "M 1.3";
//;
      A(    ;
      O     "S 2.0";
      O     "M 171.5";
      )     ;
      R     "M 1.3";
NETWORK
TITLE =Door Open Feeder - Fault

      AN    "E 12.5";
      S     "M 1.5";
//;
      A(    ;
      O     "S 2.7";
      O     "M 0.2";
      O     "M 171.5";
      )     ;
      A     "E 12.5";
      R     "M 1.5";
NETWORK
TITLE =Door Open Elevator - Fault

      AN    "E 4.6";
      S     "M 1.6";
//;
      A(    ;
      O     "S 4.7";
      O     "M 0.2";
      O     "M 171.5";
      )     ;
      A     "E 4.6";
      R     "M 1.6";
NETWORK
TITLE =Door Open Flipper - Fault
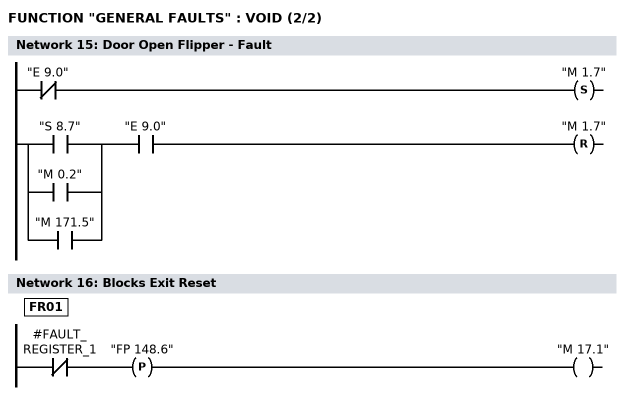

      AN    "E 9.0";
      S     "M 1.7";
//;
      A(    ;
      O     "S 8.7";
      O     "M 0.2";
      O     "M 171.5";
      )     ;
      A     "E 9.0";
      R     "M 1.7";
NETWORK
TITLE =Blocks Exit Reset

FR01: NOP   0;

      AN    #FAULT_REGISTER_1;
      FP    "FP 148.6";
      =     "M 17.1";
NETWORK
TITLE =Faults Register 2 - Conveyor 0 to Conveyor 3

      A(    ;
      L     "MB 2";
      L     0;
      <>I   ;
      )     ;
      =     #FAULT_REGISTER_2;
      =     "HMI_DB".SCREEN_CALL_1;
//;
      A     #FAULT_REGISTER_2;
      O     #CHECK_PULSE;
      O     "M 17.2";
      O     "M 9.1";
      JNB   FR02;
NETWORK
TITLE =K62.0 / 1 Conveyor 0 - Fault
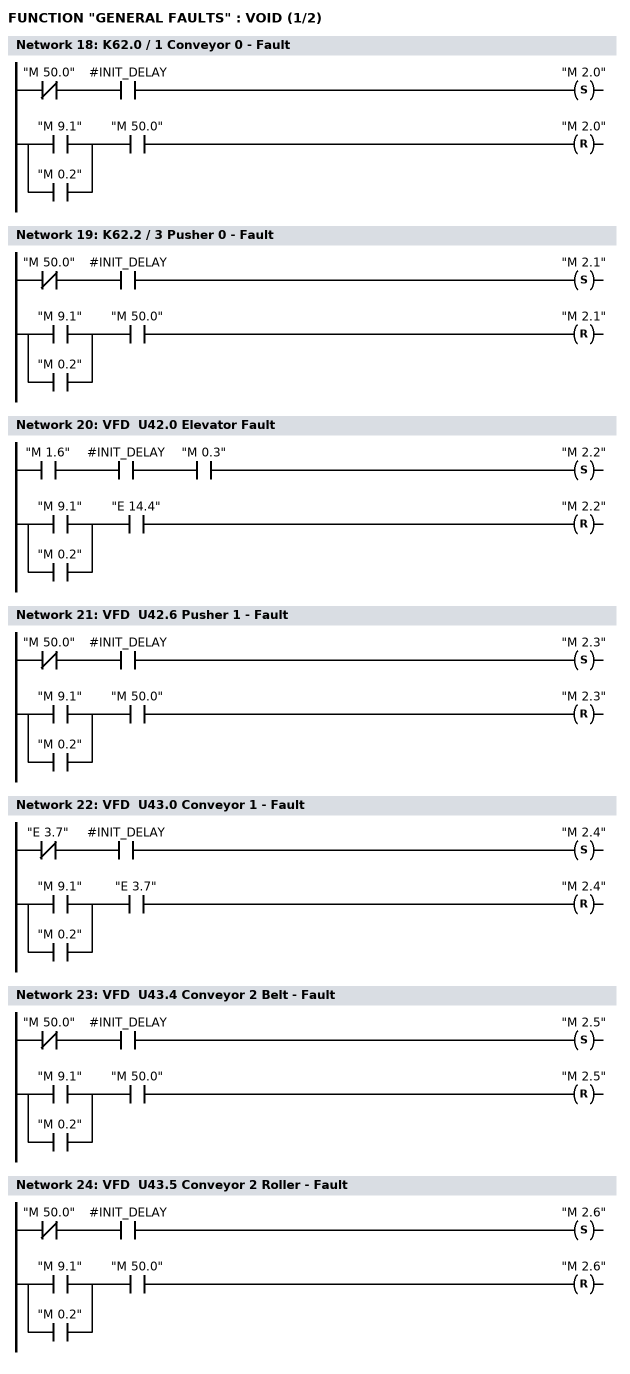

      AN    "M 50.0";
      A     #INIT_DELAY;
      S     "M 2.0";
//;
      A(    ;
      O     "M 9.1";
      O     "M 0.2";
      )     ;
      A     "M 50.0";
      R     "M 2.0";
NETWORK
TITLE =K62.2 / 3 Pusher 0 - Fault

      AN    "M 50.0";
      A     #INIT_DELAY;
      S     "M 2.1";
//;
      A(    ;
      O     "M 9.1";
      O     "M 0.2";
      )     ;
      A     "M 50.0";
      R     "M 2.1";
NETWORK
TITLE =VFD  U42.0 Elevator Fault

//   AN    #ELEVATOR_U42_0
      A     "M 1.6";
      A     #INIT_DELAY;
      A     "M 0.3";
      S     "M 2.2";
//;
      A(    ;
      O     "M 9.1";
      O     "M 0.2";
      )     ;
//      A     "E 3.6"
      A     "E 14.4";
      R     "M 2.2";
NETWORK
TITLE =VFD  U42.6 Pusher 1 - Fault

      AN    "M 50.0";
      A     #INIT_DELAY;
      S     "M 2.3";
//;
      A(    ;
      O     "M 9.1";
      O     "M 0.2";
      )     ;
      A     "M 50.0";
      R     "M 2.3";
NETWORK
TITLE =VFD  U43.0 Conveyor 1 - Fault

      AN    "E 3.7";
      A     #INIT_DELAY;
      S     "M 2.4";
//;
      A(    ;
      O     "M 9.1";
      O     "M 0.2";
      )     ;
      A     "E 3.7";
      R     "M 2.4";
NETWORK
TITLE =VFD  U43.4 Conveyor 2 Belt - Fault

      AN    "M 50.0";
      A     #INIT_DELAY;
      S     "M 2.5";
//;
      A(    ;
      O     "M 9.1";
      O     "M 0.2";
      )     ;
      A     "M 50.0";
      R     "M 2.5";
NETWORK
TITLE =VFD  U43.5 Conveyor 2 Roller - Fault

      AN    "M 50.0";
      A     #INIT_DELAY;
      S     "M 2.6";
//;
      A(    ;
      O     "M 9.1";
      O     "M 0.2";
      )     ;
      A     "M 50.0";
      R     "M 2.6";
NETWORK
TITLE =VFD  U44.0 Conveyor 3 Fault
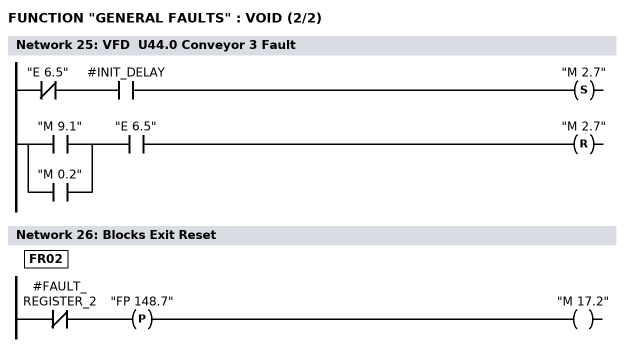

      AN    "E 6.5";
      A     #INIT_DELAY;
      S     "M 2.7";
//;
      A(    ;
      O     "M 9.1";
      O     "M 0.2";
      )     ;
      A     "E 6.5";
      R     "M 2.7";
NETWORK
TITLE =Blocks Exit Reset

FR02: NOP   0;

      AN    #FAULT_REGISTER_2;
      FP    "FP 148.7";
      =     "M 17.2";
NETWORK
TITLE =Faults Register 3 - Conveyor 4 to Conveyor 9

      A(    ;
      L     "MB 3";
      L     0;
      <>I   ;
      )     ;
      =     #FAULT_REGISTER_3;
      =     "HMI_DB".SCREEN_CALL_2;
//;
      A     #FAULT_REGISTER_3;
      O     #CHECK_PULSE;
      O     "M 17.3";
      O     "M 9.1";
      JNB   FR03;
NETWORK
TITLE =VFD  U44.3 Fault
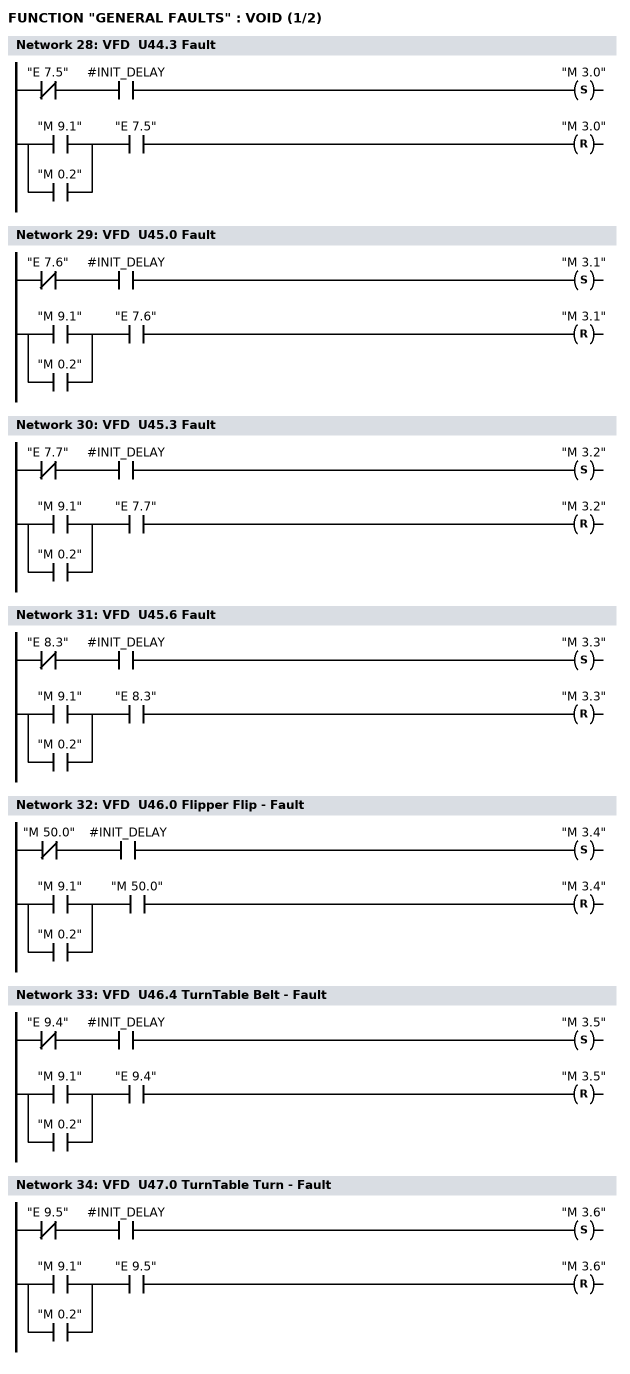

      AN    "E 7.5";
      A     #INIT_DELAY;
      S     "M 3.0";
//;
      A(    ;
      O     "M 9.1";
      O     "M 0.2";
      )     ;
      A     "E 7.5";
      R     "M 3.0";
NETWORK
TITLE =VFD  U45.0 Fault

      AN    "E 7.6";
      A     #INIT_DELAY;
      S     "M 3.1";
//;
      A(    ;
      O     "M 9.1";
      O     "M 0.2";
      )     ;
      A     "E 7.6";
      R     "M 3.1";
NETWORK
TITLE =VFD  U45.3 Fault

      AN    "E 7.7";
      A     #INIT_DELAY;
      S     "M 3.2";
//;
      A(    ;
      O     "M 9.1";
      O     "M 0.2";
      )     ;
      A     "E 7.7";
      R     "M 3.2";
NETWORK
TITLE =VFD  U45.6 Fault

      AN    "E 8.3";
      A     #INIT_DELAY;
      S     "M 3.3";
///;
      A(    ;
      O     "M 9.1";
      O     "M 0.2";
      )     ;
      A     "E 8.3";
      R     "M 3.3";
NETWORK
TITLE =VFD  U46.0 Flipper Flip - Fault

      AN    "M 50.0";
      A     #INIT_DELAY;
      S     "M 3.4";
//;
      A(    ;
      O     "M 9.1";
      O     "M 0.2";
      )     ;
      A     "M 50.0";
      R     "M 3.4";
NETWORK
TITLE =VFD  U46.4 TurnTable Belt - Fault

      AN    "E 9.4";
      A     #INIT_DELAY;
      S     "M 3.5";
//;
      A(    ;
      O     "M 9.1";
      O     "M 0.2";
      )     ;
      A     "E 9.4";
      R     "M 3.5";
NETWORK
TITLE =VFD  U47.0 TurnTable Turn - Fault

      AN    "E 9.5";
      A     #INIT_DELAY;
      S     "M 3.6";
//;
      A(    ;
      O     "M 9.1";
      O     "M 0.2";
      )     ;
      A     "E 9.5";
      R     "M 3.6";
NETWORK
TITLE =VFD  U47.5 Conveyor 9 - Fault
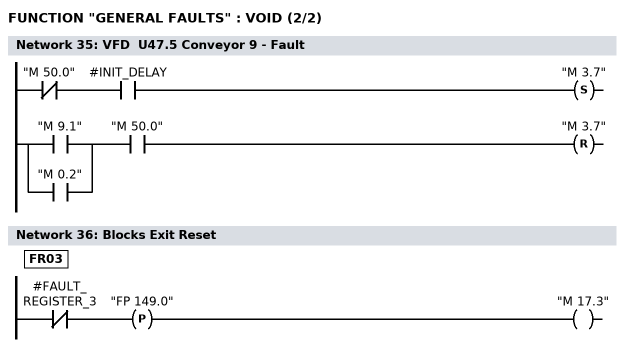

      AN    "M 50.0";
      A     #INIT_DELAY;
      S     "M 3.7";
//;
      A(    ;
      O     "M 9.1";
      O     "M 0.2";
      )     ;
      A     "M 50.0";
      R     "M 3.7";
NETWORK
TITLE =Blocks Exit Reset

FR03: NOP   0;

      AN    #FAULT_REGISTER_3;
      FP    "FP 149.0";
      =     "M 17.3";
NETWORK
TITLE =Faults Register 4 - Pusher 2 to Conveyor 23

      A(    ;
      L     "MB 4";
      L     0;
      <>I   ;
      )     ;
      =     #FAULT_REGISTER_4;
      =     "HMI_DB".SCREEN_CALL_2;
//;
      A     #FAULT_REGISTER_4;
      O     #CHECK_PULSE;
      O     "M 17.4";
      O     "M 9.1";
      JNB   FR04;
NETWORK
TITLE =VFD  U47.6 Pusher 2 - Fault
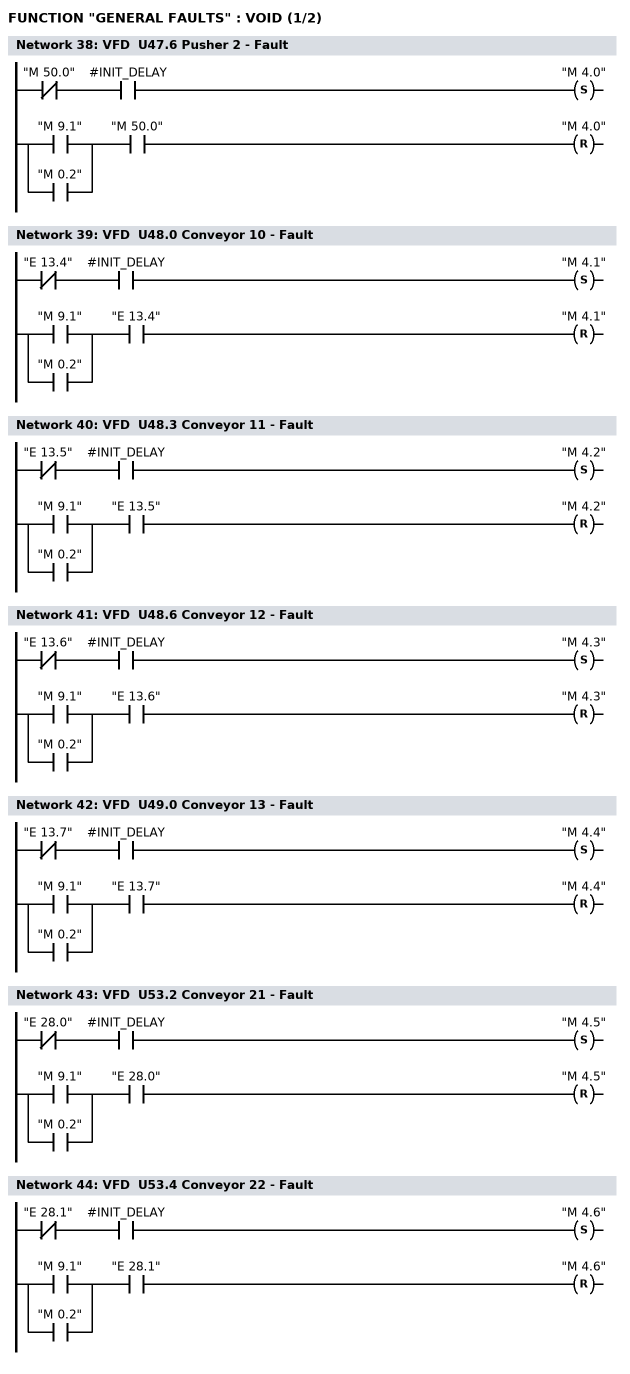

      AN    "M 50.0";
      A     #INIT_DELAY;
      S     "M 4.0";
//;
      A(    ;
      O     "M 9.1";
      O     "M 0.2";
      )     ;
      A     "M 50.0";
      R     "M 4.0";
NETWORK
TITLE =VFD  U48.0 Conveyor 10 - Fault

      AN    "E 13.4";
      A     #INIT_DELAY;
      S     "M 4.1";
//;
      A(    ;
      O     "M 9.1";
      O     "M 0.2";
      )     ;
      A     "E 13.4";
      R     "M 4.1";
NETWORK
TITLE =VFD  U48.3 Conveyor 11 - Fault

      AN    "E 13.5";
      A     #INIT_DELAY;
      S     "M 4.2";
//;
      A(    ;
      O     "M 9.1";
      O     "M 0.2";
      )     ;
      A     "E 13.5";
      R     "M 4.2";
NETWORK
TITLE =VFD  U48.6 Conveyor 12 - Fault

      AN    "E 13.6";
      A     #INIT_DELAY;
      S     "M 4.3";
//;
      A(    ;
      O     "M 9.1";
      O     "M 0.2";
      )     ;
      A     "E 13.6";
      R     "M 4.3";
NETWORK
TITLE =VFD  U49.0 Conveyor 13 - Fault

      AN    "E 13.7";
      A     #INIT_DELAY;
      S     "M 4.4";
//;
      A(    ;
      O     "M 9.1";
      O     "M 0.2";
      )     ;
      A     "E 13.7";
      R     "M 4.4";
NETWORK
TITLE =VFD  U53.2 Conveyor 21 - Fault

      AN    "E 28.0";
      A     #INIT_DELAY;
      S     "M 4.5";
//;
      A(    ;
      O     "M 9.1";
      O     "M 0.2";
      )     ;
      A     "E 28.0";
      R     "M 4.5";
NETWORK
TITLE =VFD  U53.4 Conveyor 22 - Fault

      AN    "E 28.1";
      A     #INIT_DELAY;
      S     "M 4.6";
//;
      A(    ;
      O     "M 9.1";
      O     "M 0.2";
      )     ;
      A     "E 28.1";
      R     "M 4.6";
NETWORK
TITLE =VFD  U54.0 Conveyor 23 - Fault
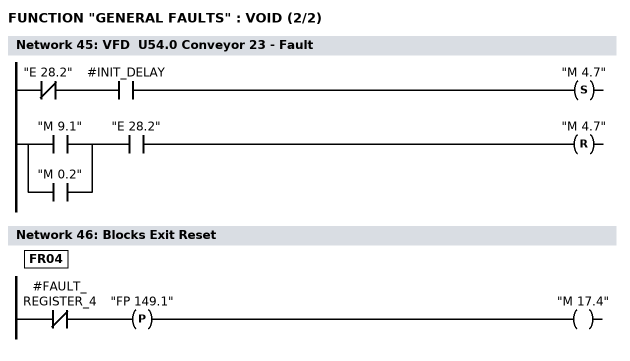

      AN    "E 28.2";
      A     #INIT_DELAY;
      S     "M 4.7";
//;
      A(    ;
      O     "M 9.1";
      O     "M 0.2";
      )     ;
      A     "E 28.2";
      R     "M 4.7";
NETWORK
TITLE =Blocks Exit Reset

FR04: NOP   0;

      AN    #FAULT_REGISTER_4;
      FP    "FP 149.1";
      =     "M 17.4";
NETWORK
TITLE =Faults Register 5 - Feeder

      A(    ;
      O     "M 7.0";
      O     "M 7.1";
      O     "M 7.2";
      )     ;
      =     #FAULT_REGISTER_5;
      =     "HMI_DB".SCREEN_CALL_3;
//;
      A     #FAULT_REGISTER_5;
      O     #CHECK_PULSE;
      O     "M 17.5";
      O     "M 9.1";
      JNB   FR05;
NETWORK
TITLE =VFD  U50.0 Feeder Lift - Fault
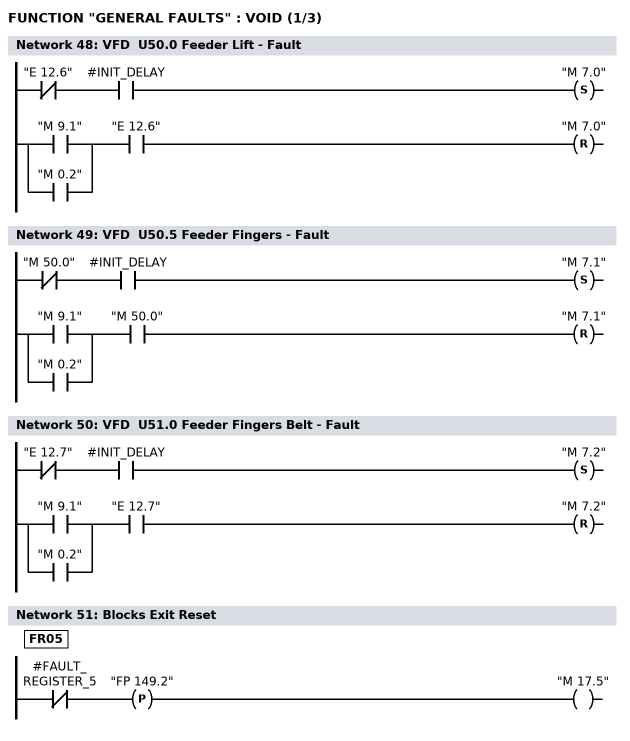

      AN    "E 12.6";
      A     #INIT_DELAY;
      S     "M 7.0";
//;
      A(    ;
      O     "M 9.1";
      O     "M 0.2";
      )     ;
      A     "E 12.6";
      R     "M 7.0";
NETWORK
TITLE =VFD  U50.5 Feeder Fingers - Fault

      AN    "M 50.0";
      A     #INIT_DELAY;
      S     "M 7.1";
//;
      A(    ;
      O     "M 9.1";
      O     "M 0.2";
      )     ;
      A     "M 50.0";
      R     "M 7.1";
NETWORK
TITLE =VFD  U51.0 Feeder Fingers Belt - Fault

      AN    "E 12.7";
      A     #INIT_DELAY;
      S     "M 7.2";
//;
      A(    ;
      O     "M 9.1";
      O     "M 0.2";
      )     ;
      A     "E 12.7";
      R     "M 7.2";
NETWORK
TITLE =Blocks Exit Reset

FR05: NOP   0;

      AN    #FAULT_REGISTER_5;
      FP    "FP 149.2";
      =     "M 17.5";
NETWORK
TITLE =Fault Status Lamp X120
